// TIA Portal V20 export
// export: Created 2026-10-20T12:39:30.7163103Z, ExportSetting WithDefaults, DisplayName Totally Integrated Automation Portal, DisplayVersion V20 Update 6, DisplayName TIA Portal Openness, DisplayVersion V20 Update 6, DisplayName TIA Portal Version Control Interface, DisplayVersion V20 Update 6, DisplayName SINAMICS Startdrive Advanced, DisplayVersion V20 SP1, DisplayName SINAMICS Startdrive G130, G150, S120, S150, SINAMICS MV, G220, S200, S210, DisplayVersion V20 SP1, DisplayName SINAMICS Startdrive G110M, G120, G120C, G120D, G120P, G115D, DisplayVersion V20 SP1, DisplayName STEP 7 Professional, DisplayVersion V20 Update 6, DisplayName STEP 7 Safety, DisplayVersion V20 Update 2, DisplayName WinCC Basic/Comfort/Advanced, DisplayVersion V20 Update 6, DisplayName WinCC Unified, DisplayVersion V20 Update 6
ORGANIZATION_BLOCK "Main"   // OB1, LAD, ProgramCycle
TITLE = "Main Program Sweep (Cycle)"
{ S7_Optimized_Access := 'TRUE' }
VERSION : 0.1
// stored: AutoNumber true, IsIECCheckEnabled false, SetENOAutomatically false
   VAR_INPUT
      Initial_Call : Bool;   // Initial call of this OB
      Remanence : Bool;   // =True, if remanent data are available
   END_VAR
   VAR_TEMP
      Fault_Handshake_Infeed_1 : Bool;
      Fault_Handshake_Outfeed_1 : Bool;
      Fault_Handshake_Infeed_2 : Bool;
      Fault_Handshake_Infeed_3 : Bool;
      Fault_Handshake_Outfeed_2 : Bool;
      Fault_Handshake_Outfeed_3 : Bool;
   END_VAR
   VAR_TEMP   // added for the SCL form of the ladder/FBD networks
      _w1 : Bool;
      _w2 : Bool;
      _w3 : Bool;
      _w4 : Bool;
      _w5 : Bool;
      _w6 : Bool;
      _w7 : Bool;
      _w8 : Bool;
      _w9 : Bool;
      _w10 : Bool;
      _w11 : Bool;
      _w12 : Bool;
      _w13 : Bool;
      _w14 : Bool;
      _w15 : Bool;
   END_VAR
BEGIN

REGION Network 1: START PLC
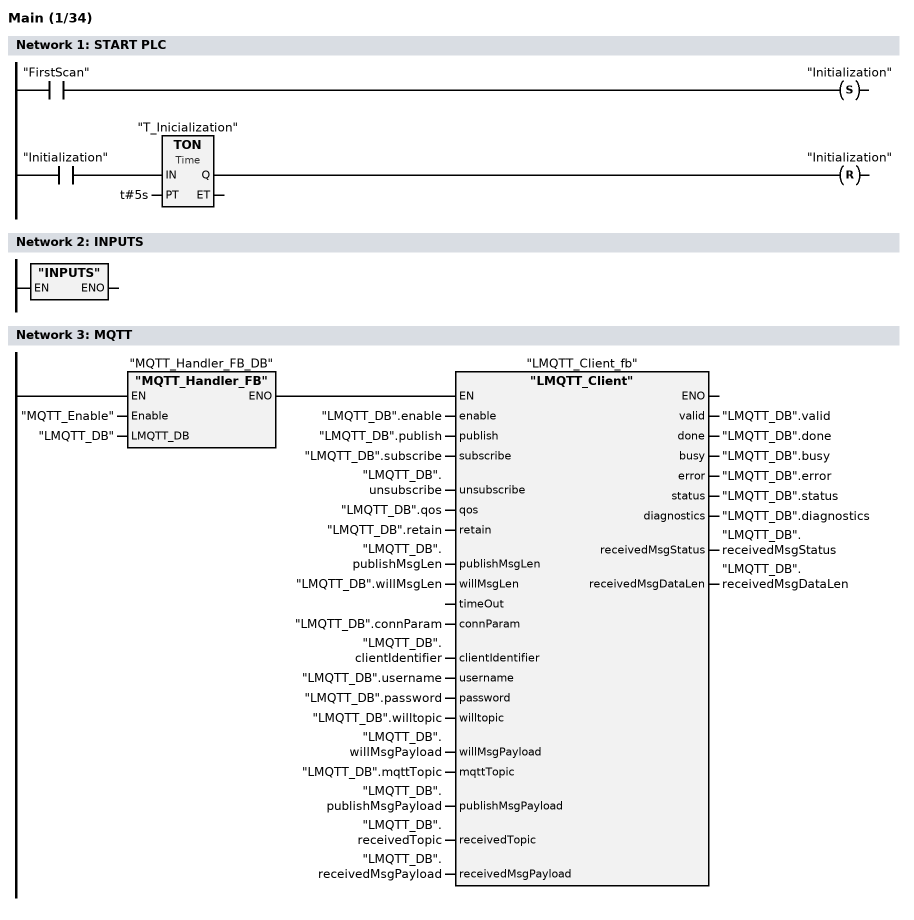
   RUNG wire#powerrail
      Contact( "FirstScan" )
      S_Coil( "Initialization" )
   END_RUNG
   RUNG wire#powerrail
      Contact( "Initialization" )
      { S7_Templates := "time_type := Time" } "T_Inicialization".TON(pt := t#5s, et =>)
      R_Coil( "Initialization" )
   END_RUNG
   // the same network as SCL:
   IF "FirstScan" THEN "Initialization" := TRUE; END_IF;
   "T_Inicialization".TON(IN := "Initialization", PT := t#5s);
   IF "T_Inicialization".Q THEN "Initialization" := FALSE; END_IF;
END_REGION

REGION Network 2: INPUTS
   RUNG wire#powerrail
      "INPUTS"()
   END_RUNG
   // the same network as SCL:
   "INPUTS"();
END_REGION

REGION Network 3: MQTT
   RUNG wire#powerrail
      "MQTT_Handler_FB_DB"(Enable := "MQTT_Enable", LMQTT_DB := "LMQTT_DB")
      "LMQTT_Client_fb"(enable := "LMQTT_DB".enable, publish := "LMQTT_DB".publish, subscribe := "LMQTT_DB".subscribe, unsubscribe := "LMQTT_DB".unsubscribe, qos := "LMQTT_DB".qos, retain := "LMQTT_DB".retain, publishMsgLen := "LMQTT_DB".publishMsgLen, willMsgLen := "LMQTT_DB".willMsgLen, timeOut :=, connParam := "LMQTT_DB".connParam, clientIdentifier := "LMQTT_DB".clientIdentifier, username := "LMQTT_DB".username, password := "LMQTT_DB".password, willtopic := "LMQTT_DB".willtopic, willMsgPayload := "LMQTT_DB".willMsgPayload, mqttTopic := "LMQTT_DB".mqttTopic, publishMsgPayload := "LMQTT_DB".publishMsgPayload, receivedTopic := "LMQTT_DB".receivedTopic, receivedMsgPayload := "LMQTT_DB".receivedMsgPayload, valid => "LMQTT_DB".valid, done => "LMQTT_DB".done, busy => "LMQTT_DB".busy, error => "LMQTT_DB".error, status => "LMQTT_DB".status, diagnostics => "LMQTT_DB".diagnostics, receivedMsgStatus => "LMQTT_DB".receivedMsgStatus, receivedMsgDataLen => "LMQTT_DB".receivedMsgDataLen)
   END_RUNG
   // the same network as SCL:
   "MQTT_Handler_FB_DB"(Enable := "MQTT_Enable", LMQTT_DB := "LMQTT_DB", ENO => #_w1);   // "MQTT_Handler_FB"
   IF #_w1 THEN
       "LMQTT_Client_fb"(enable := "LMQTT_DB".enable,   // "LMQTT_Client"
                         publish := "LMQTT_DB".publish,
                         subscribe := "LMQTT_DB".subscribe,
                         unsubscribe := "LMQTT_DB".unsubscribe,
                         qos := "LMQTT_DB".qos,
                         retain := "LMQTT_DB".retain,
                         publishMsgLen := "LMQTT_DB".publishMsgLen,
                         willMsgLen := "LMQTT_DB".willMsgLen,
                         connParam := "LMQTT_DB".connParam,
                         clientIdentifier := "LMQTT_DB".clientIdentifier,
                         username := "LMQTT_DB".username,
                         password := "LMQTT_DB".password,
                         willtopic := "LMQTT_DB".willtopic,
                         willMsgPayload := "LMQTT_DB".willMsgPayload,
                         mqttTopic := "LMQTT_DB".mqttTopic,
                         publishMsgPayload := "LMQTT_DB".publishMsgPayload,
                         receivedTopic := "LMQTT_DB".receivedTopic,
                         receivedMsgPayload := "LMQTT_DB".receivedMsgPayload,
                         valid => "LMQTT_DB".valid,
                         done => "LMQTT_DB".done,
                         busy => "LMQTT_DB".busy,
                         error => "LMQTT_DB".error,
                         status => "LMQTT_DB".status,
                         diagnostics => "LMQTT_DB".diagnostics,
                         receivedMsgStatus => "LMQTT_DB".receivedMsgStatus,
                         receivedMsgDataLen => "LMQTT_DB".receivedMsgDataLen);
   END_IF;
END_REGION

REGION Network 4: Absolute Encoders
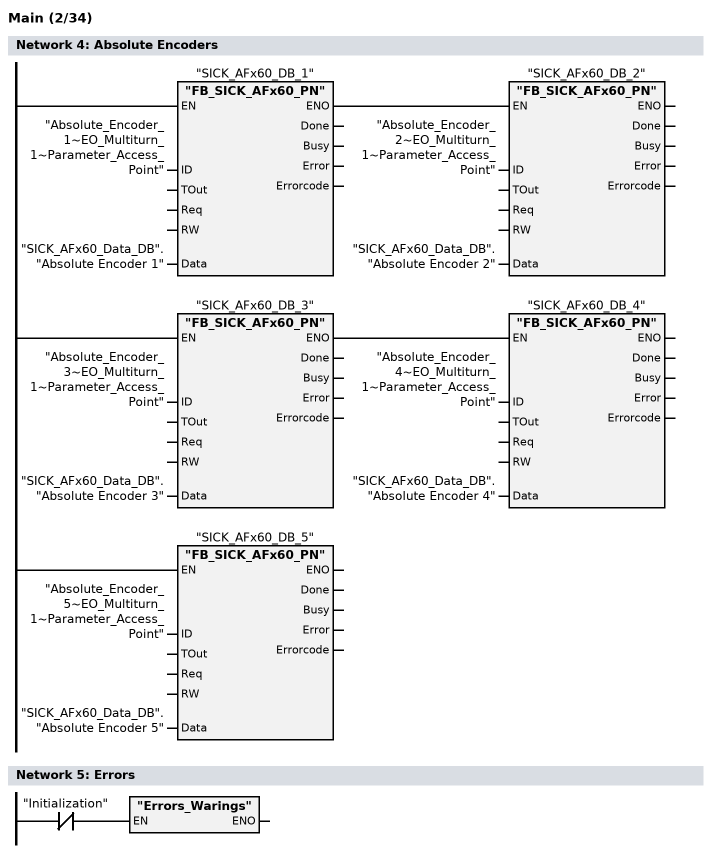
   RUNG wire#powerrail
      "SICK_AFx60_DB_1"(ID := "Absolute_Encoder_1~EO_Multiturn_1~Parameter_Access_Point", TOut :=, Req :=, RW :=, Data := "SICK_AFx60_Data_DB"."Absolute Encoder 1", Done =>, Busy =>, Error =>, Errorcode =>)
      "SICK_AFx60_DB_2"(ID := "Absolute_Encoder_2~EO_Multiturn_1~Parameter_Access_Point", TOut :=, Req :=, RW :=, Data := "SICK_AFx60_Data_DB"."Absolute Encoder 2", Done =>, Busy =>, Error =>, Errorcode =>)
   END_RUNG
   RUNG wire#powerrail
      "SICK_AFx60_DB_3"(ID := "Absolute_Encoder_3~EO_Multiturn_1~Parameter_Access_Point", TOut :=, Req :=, RW :=, Data := "SICK_AFx60_Data_DB"."Absolute Encoder 3", Done =>, Busy =>, Error =>, Errorcode =>)
      "SICK_AFx60_DB_4"(ID := "Absolute_Encoder_4~EO_Multiturn_1~Parameter_Access_Point", TOut :=, Req :=, RW :=, Data := "SICK_AFx60_Data_DB"."Absolute Encoder 4", Done =>, Busy =>, Error =>, Errorcode =>)
   END_RUNG
   RUNG wire#powerrail
      "SICK_AFx60_DB_5"(ID := "Absolute_Encoder_5~EO_Multiturn_1~Parameter_Access_Point", TOut :=, Req :=, RW :=, Data := "SICK_AFx60_Data_DB"."Absolute Encoder 5", Done =>, Busy =>, Error =>, Errorcode =>)
   END_RUNG
   // the same network as SCL:
   "SICK_AFx60_DB_1"(ID := "Absolute_Encoder_1~EO_Multiturn_1~Parameter_Access_Point",   // "FB_SICK_AFx60_PN"
                     Data := "SICK_AFx60_Data_DB"."Absolute Encoder 1",
                     ENO => #_w1);
   IF #_w1 THEN
       "SICK_AFx60_DB_2"(ID := "Absolute_Encoder_2~EO_Multiturn_1~Parameter_Access_Point",   // "FB_SICK_AFx60_PN"
                         Data := "SICK_AFx60_Data_DB"."Absolute Encoder 2");
   END_IF;
   "SICK_AFx60_DB_3"(ID := "Absolute_Encoder_3~EO_Multiturn_1~Parameter_Access_Point",   // "FB_SICK_AFx60_PN"
                     Data := "SICK_AFx60_Data_DB"."Absolute Encoder 3",
                     ENO => #_w2);
   IF #_w2 THEN
       "SICK_AFx60_DB_4"(ID := "Absolute_Encoder_4~EO_Multiturn_1~Parameter_Access_Point",   // "FB_SICK_AFx60_PN"
                         Data := "SICK_AFx60_Data_DB"."Absolute Encoder 4");
   END_IF;
   "SICK_AFx60_DB_5"(ID := "Absolute_Encoder_5~EO_Multiturn_1~Parameter_Access_Point",   // "FB_SICK_AFx60_PN"
                     Data := "SICK_AFx60_Data_DB"."Absolute Encoder 5");
END_REGION

REGION Network 5: Errors
   RUNG wire#powerrail
      I_Contact( "Initialization" )
      "Errors_Warings"()
   END_RUNG
   // the same network as SCL:
   IF NOT "Initialization" THEN "Errors_Warings"(); END_IF;
END_REGION

REGION Network 6: AUTO TEST 1
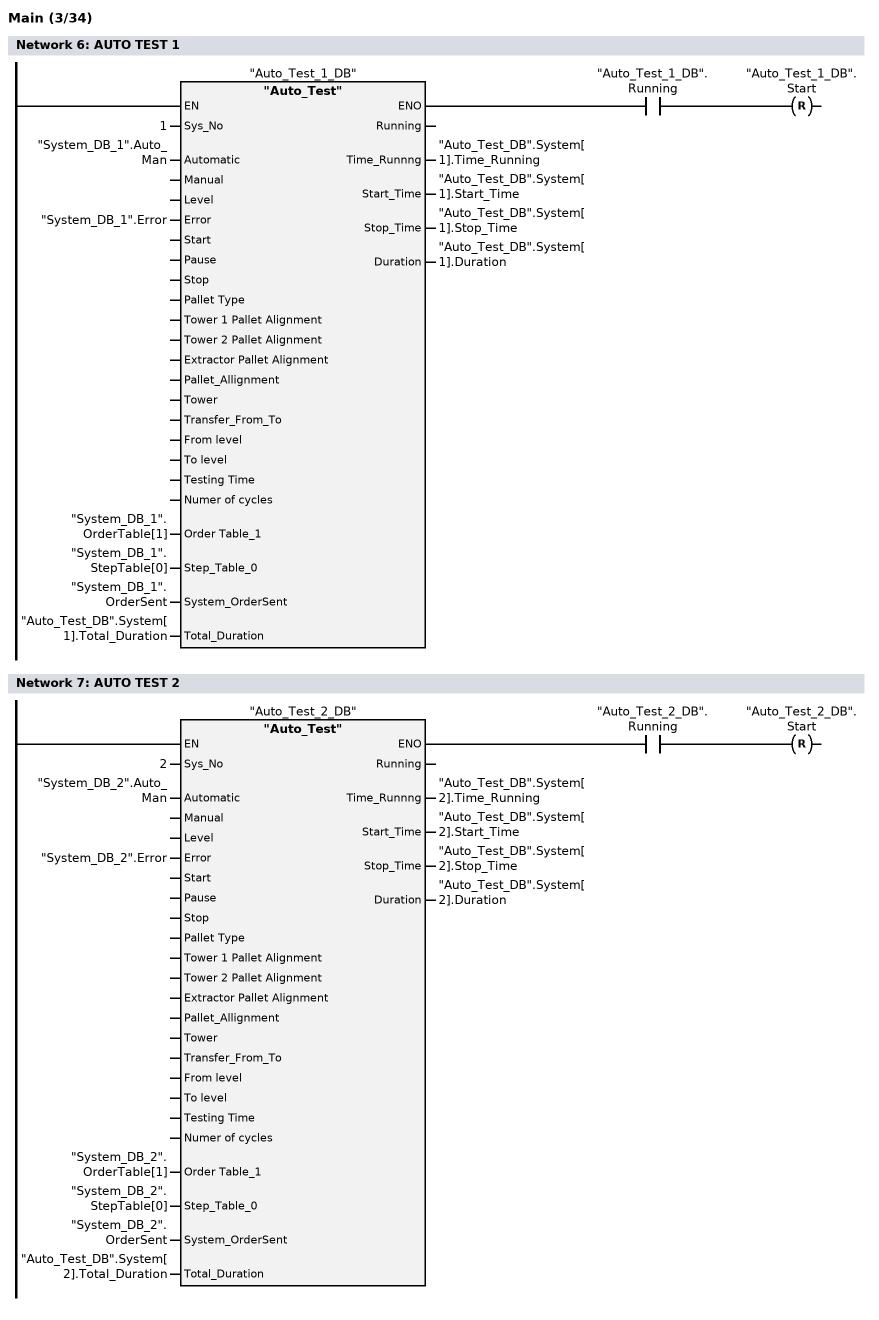
   RUNG wire#powerrail
      "Auto_Test_1_DB"(Sys_No := 1, Automatic := "System_DB_1".Auto_Man, Manual :=, Level :=, Error := "System_DB_1".Error, Start :=, Pause :=, Stop :=, "Pallet Type" :=, "Tower 1 Pallet Alignment" :=, "Tower 2 Pallet Alignment" :=, "Extractor Pallet Alignment" :=, Pallet_Allignment :=, Tower :=, Transfer_From_To :=, "From level" :=, "To level" :=, "Testing Time" :=, "Numer of cycles" :=, "Order Table_1" := "System_DB_1".OrderTable[1], Step_Table_0 := "System_DB_1".StepTable[0], System_OrderSent := "System_DB_1".OrderSent, Total_Duration := "Auto_Test_DB".System[1].Total_Duration, Running =>, Time_Runnng => "Auto_Test_DB".System[1].Time_Running, Start_Time => "Auto_Test_DB".System[1].Start_Time, Stop_Time => "Auto_Test_DB".System[1].Stop_Time, Duration => "Auto_Test_DB".System[1].Duration)
      Contact( "Auto_Test_1_DB".Running )
      R_Coil( "Auto_Test_1_DB".Start )
   END_RUNG
   // the same network as SCL:
   "Auto_Test_1_DB"(Sys_No := 1,   // "Auto_Test"
                    Automatic := "System_DB_1".Auto_Man,
                    Error := "System_DB_1".Error,
                    "Order Table_1" := "System_DB_1".OrderTable[1],
                    Step_Table_0 := "System_DB_1".StepTable[0],
                    System_OrderSent := "System_DB_1".OrderSent,
                    Total_Duration := "Auto_Test_DB".System[1].Total_Duration,
                    Time_Runnng => "Auto_Test_DB".System[1].Time_Running,
                    Start_Time => "Auto_Test_DB".System[1].Start_Time,
                    Stop_Time => "Auto_Test_DB".System[1].Stop_Time,
                    Duration => "Auto_Test_DB".System[1].Duration,
                    ENO => #_w1);
   IF #_w1 AND "Auto_Test_1_DB".Running THEN "Auto_Test_1_DB".Start := FALSE; END_IF;
END_REGION

REGION Network 7: AUTO TEST 2
   RUNG wire#powerrail
      "Auto_Test_2_DB"(Sys_No := 2, Automatic := "System_DB_2".Auto_Man, Manual :=, Level :=, Error := "System_DB_2".Error, Start :=, Pause :=, Stop :=, "Pallet Type" :=, "Tower 1 Pallet Alignment" :=, "Tower 2 Pallet Alignment" :=, "Extractor Pallet Alignment" :=, Pallet_Allignment :=, Tower :=, Transfer_From_To :=, "From level" :=, "To level" :=, "Testing Time" :=, "Numer of cycles" :=, "Order Table_1" := "System_DB_2".OrderTable[1], Step_Table_0 := "System_DB_2".StepTable[0], System_OrderSent := "System_DB_2".OrderSent, Total_Duration := "Auto_Test_DB".System[2].Total_Duration, Running =>, Time_Runnng => "Auto_Test_DB".System[2].Time_Running, Start_Time => "Auto_Test_DB".System[2].Start_Time, Stop_Time => "Auto_Test_DB".System[2].Stop_Time, Duration => "Auto_Test_DB".System[2].Duration)
      Contact( "Auto_Test_2_DB".Running )
      R_Coil( "Auto_Test_2_DB".Start )
   END_RUNG
   // the same network as SCL:
   "Auto_Test_2_DB"(Sys_No := 2,   // "Auto_Test"
                    Automatic := "System_DB_2".Auto_Man,
                    Error := "System_DB_2".Error,
                    "Order Table_1" := "System_DB_2".OrderTable[1],
                    Step_Table_0 := "System_DB_2".StepTable[0],
                    System_OrderSent := "System_DB_2".OrderSent,
                    Total_Duration := "Auto_Test_DB".System[2].Total_Duration,
                    Time_Runnng => "Auto_Test_DB".System[2].Time_Running,
                    Start_Time => "Auto_Test_DB".System[2].Start_Time,
                    Stop_Time => "Auto_Test_DB".System[2].Stop_Time,
                    Duration => "Auto_Test_DB".System[2].Duration,
                    ENO => #_w1);
   IF #_w1 AND "Auto_Test_2_DB".Running THEN "Auto_Test_2_DB".Start := FALSE; END_IF;
END_REGION

REGION Network 8: AUTO TEST 3
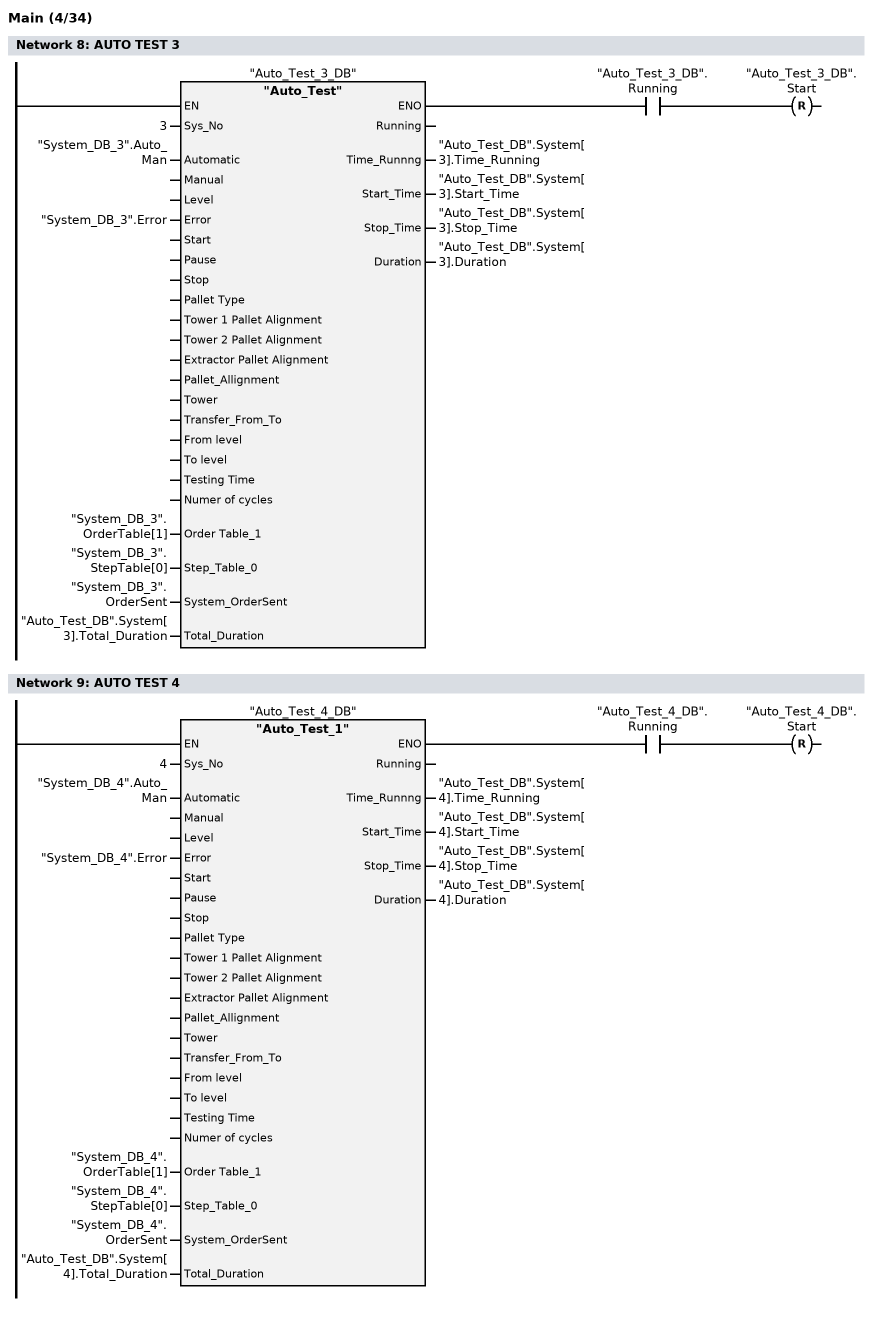
   RUNG wire#powerrail
      "Auto_Test_3_DB"(Sys_No := 3, Automatic := "System_DB_3".Auto_Man, Manual :=, Level :=, Error := "System_DB_3".Error, Start :=, Pause :=, Stop :=, "Pallet Type" :=, "Tower 1 Pallet Alignment" :=, "Tower 2 Pallet Alignment" :=, "Extractor Pallet Alignment" :=, Pallet_Allignment :=, Tower :=, Transfer_From_To :=, "From level" :=, "To level" :=, "Testing Time" :=, "Numer of cycles" :=, "Order Table_1" := "System_DB_3".OrderTable[1], Step_Table_0 := "System_DB_3".StepTable[0], System_OrderSent := "System_DB_3".OrderSent, Total_Duration := "Auto_Test_DB".System[3].Total_Duration, Running =>, Time_Runnng => "Auto_Test_DB".System[3].Time_Running, Start_Time => "Auto_Test_DB".System[3].Start_Time, Stop_Time => "Auto_Test_DB".System[3].Stop_Time, Duration => "Auto_Test_DB".System[3].Duration)
      Contact( "Auto_Test_3_DB".Running )
      R_Coil( "Auto_Test_3_DB".Start )
   END_RUNG
   // the same network as SCL:
   "Auto_Test_3_DB"(Sys_No := 3,   // "Auto_Test"
                    Automatic := "System_DB_3".Auto_Man,
                    Error := "System_DB_3".Error,
                    "Order Table_1" := "System_DB_3".OrderTable[1],
                    Step_Table_0 := "System_DB_3".StepTable[0],
                    System_OrderSent := "System_DB_3".OrderSent,
                    Total_Duration := "Auto_Test_DB".System[3].Total_Duration,
                    Time_Runnng => "Auto_Test_DB".System[3].Time_Running,
                    Start_Time => "Auto_Test_DB".System[3].Start_Time,
                    Stop_Time => "Auto_Test_DB".System[3].Stop_Time,
                    Duration => "Auto_Test_DB".System[3].Duration,
                    ENO => #_w1);
   IF #_w1 AND "Auto_Test_3_DB".Running THEN "Auto_Test_3_DB".Start := FALSE; END_IF;
END_REGION

REGION Network 9: AUTO TEST 4
   RUNG wire#powerrail
      "Auto_Test_4_DB"(Sys_No := 4, Automatic := "System_DB_4".Auto_Man, Manual :=, Level :=, Error := "System_DB_4".Error, Start :=, Pause :=, Stop :=, "Pallet Type" :=, "Tower 1 Pallet Alignment" :=, "Tower 2 Pallet Alignment" :=, "Extractor Pallet Alignment" :=, Pallet_Allignment :=, Tower :=, Transfer_From_To :=, "From level" :=, "To level" :=, "Testing Time" :=, "Numer of cycles" :=, "Order Table_1" := "System_DB_4".OrderTable[1], Step_Table_0 := "System_DB_4".StepTable[0], System_OrderSent := "System_DB_4".OrderSent, Total_Duration := "Auto_Test_DB".System[4].Total_Duration, Running =>, Time_Runnng => "Auto_Test_DB".System[4].Time_Running, Start_Time => "Auto_Test_DB".System[4].Start_Time, Stop_Time => "Auto_Test_DB".System[4].Stop_Time, Duration => "Auto_Test_DB".System[4].Duration)
      Contact( "Auto_Test_4_DB".Running )
      R_Coil( "Auto_Test_4_DB".Start )
   END_RUNG
   // the same network as SCL:
   "Auto_Test_4_DB"(Sys_No := 4,   // "Auto_Test_1"
                    Automatic := "System_DB_4".Auto_Man,
                    Error := "System_DB_4".Error,
                    "Order Table_1" := "System_DB_4".OrderTable[1],
                    Step_Table_0 := "System_DB_4".StepTable[0],
                    System_OrderSent := "System_DB_4".OrderSent,
                    Total_Duration := "Auto_Test_DB".System[4].Total_Duration,
                    Time_Runnng => "Auto_Test_DB".System[4].Time_Running,
                    Start_Time => "Auto_Test_DB".System[4].Start_Time,
                    Stop_Time => "Auto_Test_DB".System[4].Stop_Time,
                    Duration => "Auto_Test_DB".System[4].Duration,
                    ENO => #_w1);
   IF #_w1 AND "Auto_Test_4_DB".Running THEN "Auto_Test_4_DB".Start := FALSE; END_IF;
END_REGION

REGION Network 10: AUTO TEST 5
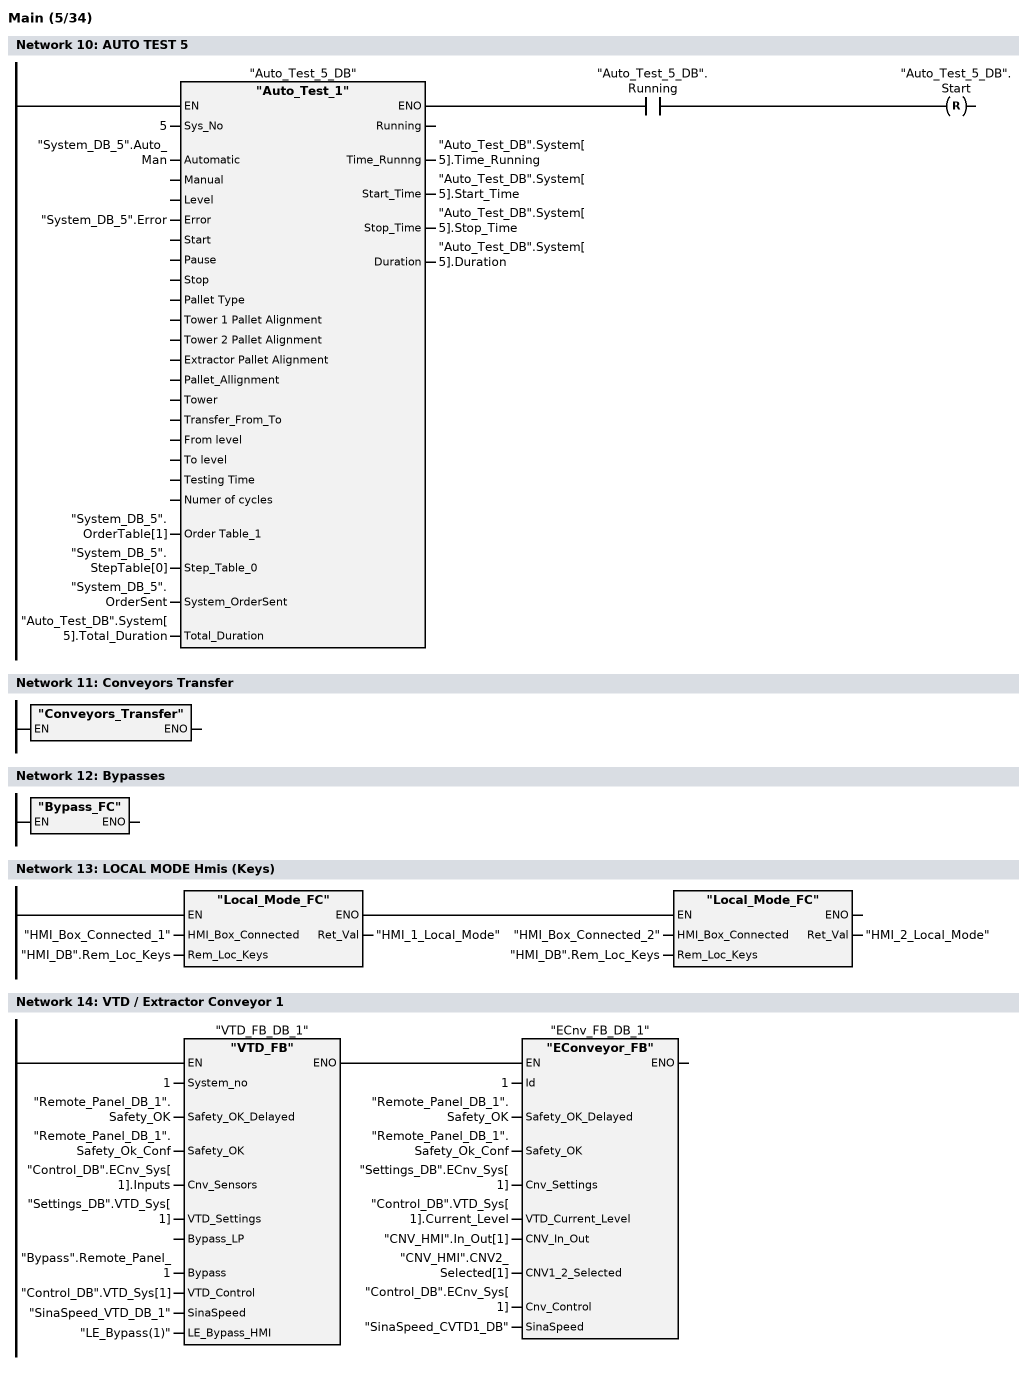
   RUNG wire#powerrail
      "Auto_Test_5_DB"(Sys_No := 5, Automatic := "System_DB_5".Auto_Man, Manual :=, Level :=, Error := "System_DB_5".Error, Start :=, Pause :=, Stop :=, "Pallet Type" :=, "Tower 1 Pallet Alignment" :=, "Tower 2 Pallet Alignment" :=, "Extractor Pallet Alignment" :=, Pallet_Allignment :=, Tower :=, Transfer_From_To :=, "From level" :=, "To level" :=, "Testing Time" :=, "Numer of cycles" :=, "Order Table_1" := "System_DB_5".OrderTable[1], Step_Table_0 := "System_DB_5".StepTable[0], System_OrderSent := "System_DB_5".OrderSent, Total_Duration := "Auto_Test_DB".System[5].Total_Duration, Running =>, Time_Runnng => "Auto_Test_DB".System[5].Time_Running, Start_Time => "Auto_Test_DB".System[5].Start_Time, Stop_Time => "Auto_Test_DB".System[5].Stop_Time, Duration => "Auto_Test_DB".System[5].Duration)
      Contact( "Auto_Test_5_DB".Running )
      R_Coil( "Auto_Test_5_DB".Start )
   END_RUNG
   // the same network as SCL:
   "Auto_Test_5_DB"(Sys_No := 5,   // "Auto_Test_1"
                    Automatic := "System_DB_5".Auto_Man,
                    Error := "System_DB_5".Error,
                    "Order Table_1" := "System_DB_5".OrderTable[1],
                    Step_Table_0 := "System_DB_5".StepTable[0],
                    System_OrderSent := "System_DB_5".OrderSent,
                    Total_Duration := "Auto_Test_DB".System[5].Total_Duration,
                    Time_Runnng => "Auto_Test_DB".System[5].Time_Running,
                    Start_Time => "Auto_Test_DB".System[5].Start_Time,
                    Stop_Time => "Auto_Test_DB".System[5].Stop_Time,
                    Duration => "Auto_Test_DB".System[5].Duration,
                    ENO => #_w1);
   IF #_w1 AND "Auto_Test_5_DB".Running THEN "Auto_Test_5_DB".Start := FALSE; END_IF;
END_REGION

REGION Network 11: Conveyors Transfer
   RUNG wire#powerrail
      "Conveyors_Transfer"()
   END_RUNG
   // the same network as SCL:
   "Conveyors_Transfer"();
END_REGION

REGION Network 12: Bypasses
   RUNG wire#powerrail
      "Bypass_FC"()
   END_RUNG
   // the same network as SCL:
   "Bypass_FC"();
END_REGION

REGION Network 13: LOCAL MODE Hmis (Keys)
   RUNG wire#powerrail
      "Local_Mode_FC"(HMI_Box_Connected := "HMI_Box_Connected_1", Rem_Loc_Keys := "HMI_DB".Rem_Loc_Keys, Ret_Val => "HMI_1_Local_Mode")
      "Local_Mode_FC"(HMI_Box_Connected := "HMI_Box_Connected_2", Rem_Loc_Keys := "HMI_DB".Rem_Loc_Keys, Ret_Val => "HMI_2_Local_Mode")
   END_RUNG
   // the same network as SCL:
   "HMI_1_Local_Mode" := "Local_Mode_FC"(HMI_Box_Connected := "HMI_Box_Connected_1",
                           Rem_Loc_Keys := "HMI_DB".Rem_Loc_Keys,
                           ENO => #_w1);
   IF #_w1 THEN
       "HMI_2_Local_Mode" := "Local_Mode_FC"(HMI_Box_Connected := "HMI_Box_Connected_2",
                               Rem_Loc_Keys := "HMI_DB".Rem_Loc_Keys);
   END_IF;
END_REGION

REGION Network 14: VTD / Extractor Conveyor 1
   RUNG wire#powerrail
      "VTD_FB_DB_1"(System_no := 1, Safety_OK_Delayed := "Remote_Panel_DB_1".Safety_OK, Safety_OK := "Remote_Panel_DB_1".Safety_Ok_Conf, Cnv_Sensors := "Control_DB".ECnv_Sys[1].Inputs, VTD_Settings := "Settings_DB".VTD_Sys[1], Bypass_LP :=, Bypass := "Bypass".Remote_Panel_1, VTD_Control := "Control_DB".VTD_Sys[1], SinaSpeed := "SinaSpeed_VTD_DB_1", LE_Bypass_HMI := "LE_Bypass(1)")
      "ECnv_FB_DB_1"(Id := 1, Safety_OK_Delayed := "Remote_Panel_DB_1".Safety_OK, Safety_OK := "Remote_Panel_DB_1".Safety_Ok_Conf, Cnv_Settings := "Settings_DB".ECnv_Sys[1], VTD_Current_Level := "Control_DB".VTD_Sys[1].Current_Level, CNV_In_Out := "CNV_HMI".In_Out[1], CNV1_2_Selected := "CNV_HMI".CNV2_Selected[1], Cnv_Control := "Control_DB".ECnv_Sys[1], SinaSpeed := "SinaSpeed_CVTD1_DB")
   END_RUNG
   // the same network as SCL:
   "VTD_FB_DB_1"(System_no := 1,   // "VTD_FB"
                 Safety_OK_Delayed := "Remote_Panel_DB_1".Safety_OK,
                 Safety_OK := "Remote_Panel_DB_1".Safety_Ok_Conf,
                 Cnv_Sensors := "Control_DB".ECnv_Sys[1].Inputs,
                 VTD_Settings := "Settings_DB".VTD_Sys[1],
                 Bypass := "Bypass".Remote_Panel_1,
                 VTD_Control := "Control_DB".VTD_Sys[1],
                 SinaSpeed := "SinaSpeed_VTD_DB_1",
                 LE_Bypass_HMI := "LE_Bypass(1)",
                 ENO => #_w1);
   IF #_w1 THEN
       "ECnv_FB_DB_1"(Id := 1,   // "EConveyor_FB"
                      Safety_OK_Delayed := "Remote_Panel_DB_1".Safety_OK,
                      Safety_OK := "Remote_Panel_DB_1".Safety_Ok_Conf,
                      Cnv_Settings := "Settings_DB".ECnv_Sys[1],
                      VTD_Current_Level := "Control_DB".VTD_Sys[1].Current_Level,
                      CNV_In_Out := "CNV_HMI".In_Out[1],
                      CNV1_2_Selected := "CNV_HMI".CNV2_Selected[1],
                      Cnv_Control := "Control_DB".ECnv_Sys[1],
                      SinaSpeed := "SinaSpeed_CVTD1_DB");
   END_IF;
END_REGION

REGION Network 15: VTD / Extractor Conveyor 2
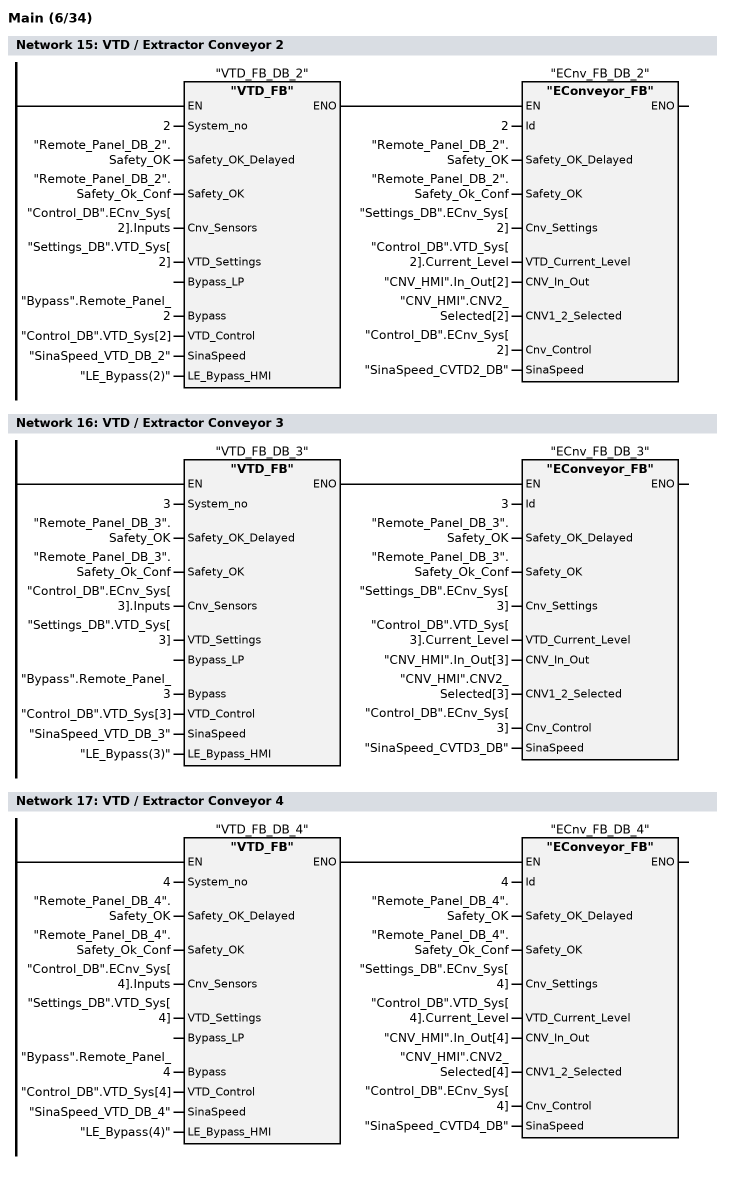
   RUNG wire#powerrail
      "VTD_FB_DB_2"(System_no := 2, Safety_OK_Delayed := "Remote_Panel_DB_2".Safety_OK, Safety_OK := "Remote_Panel_DB_2".Safety_Ok_Conf, Cnv_Sensors := "Control_DB".ECnv_Sys[2].Inputs, VTD_Settings := "Settings_DB".VTD_Sys[2], Bypass_LP :=, Bypass := "Bypass".Remote_Panel_2, VTD_Control := "Control_DB".VTD_Sys[2], SinaSpeed := "SinaSpeed_VTD_DB_2", LE_Bypass_HMI := "LE_Bypass(2)")
      "ECnv_FB_DB_2"(Id := 2, Safety_OK_Delayed := "Remote_Panel_DB_2".Safety_OK, Safety_OK := "Remote_Panel_DB_2".Safety_Ok_Conf, Cnv_Settings := "Settings_DB".ECnv_Sys[2], VTD_Current_Level := "Control_DB".VTD_Sys[2].Current_Level, CNV_In_Out := "CNV_HMI".In_Out[2], CNV1_2_Selected := "CNV_HMI".CNV2_Selected[2], Cnv_Control := "Control_DB".ECnv_Sys[2], SinaSpeed := "SinaSpeed_CVTD2_DB")
   END_RUNG
   // the same network as SCL:
   "VTD_FB_DB_2"(System_no := 2,   // "VTD_FB"
                 Safety_OK_Delayed := "Remote_Panel_DB_2".Safety_OK,
                 Safety_OK := "Remote_Panel_DB_2".Safety_Ok_Conf,
                 Cnv_Sensors := "Control_DB".ECnv_Sys[2].Inputs,
                 VTD_Settings := "Settings_DB".VTD_Sys[2],
                 Bypass := "Bypass".Remote_Panel_2,
                 VTD_Control := "Control_DB".VTD_Sys[2],
                 SinaSpeed := "SinaSpeed_VTD_DB_2",
                 LE_Bypass_HMI := "LE_Bypass(2)",
                 ENO => #_w1);
   IF #_w1 THEN
       "ECnv_FB_DB_2"(Id := 2,   // "EConveyor_FB"
                      Safety_OK_Delayed := "Remote_Panel_DB_2".Safety_OK,
                      Safety_OK := "Remote_Panel_DB_2".Safety_Ok_Conf,
                      Cnv_Settings := "Settings_DB".ECnv_Sys[2],
                      VTD_Current_Level := "Control_DB".VTD_Sys[2].Current_Level,
                      CNV_In_Out := "CNV_HMI".In_Out[2],
                      CNV1_2_Selected := "CNV_HMI".CNV2_Selected[2],
                      Cnv_Control := "Control_DB".ECnv_Sys[2],
                      SinaSpeed := "SinaSpeed_CVTD2_DB");
   END_IF;
END_REGION

REGION Network 16: VTD / Extractor Conveyor 3
   RUNG wire#powerrail
      "VTD_FB_DB_3"(System_no := 3, Safety_OK_Delayed := "Remote_Panel_DB_3".Safety_OK, Safety_OK := "Remote_Panel_DB_3".Safety_Ok_Conf, Cnv_Sensors := "Control_DB".ECnv_Sys[3].Inputs, VTD_Settings := "Settings_DB".VTD_Sys[3], Bypass_LP :=, Bypass := "Bypass".Remote_Panel_3, VTD_Control := "Control_DB".VTD_Sys[3], SinaSpeed := "SinaSpeed_VTD_DB_3", LE_Bypass_HMI := "LE_Bypass(3)")
      "ECnv_FB_DB_3"(Id := 3, Safety_OK_Delayed := "Remote_Panel_DB_3".Safety_OK, Safety_OK := "Remote_Panel_DB_3".Safety_Ok_Conf, Cnv_Settings := "Settings_DB".ECnv_Sys[3], VTD_Current_Level := "Control_DB".VTD_Sys[3].Current_Level, CNV_In_Out := "CNV_HMI".In_Out[3], CNV1_2_Selected := "CNV_HMI".CNV2_Selected[3], Cnv_Control := "Control_DB".ECnv_Sys[3], SinaSpeed := "SinaSpeed_CVTD3_DB")
   END_RUNG
   // the same network as SCL:
   "VTD_FB_DB_3"(System_no := 3,   // "VTD_FB"
                 Safety_OK_Delayed := "Remote_Panel_DB_3".Safety_OK,
                 Safety_OK := "Remote_Panel_DB_3".Safety_Ok_Conf,
                 Cnv_Sensors := "Control_DB".ECnv_Sys[3].Inputs,
                 VTD_Settings := "Settings_DB".VTD_Sys[3],
                 Bypass := "Bypass".Remote_Panel_3,
                 VTD_Control := "Control_DB".VTD_Sys[3],
                 SinaSpeed := "SinaSpeed_VTD_DB_3",
                 LE_Bypass_HMI := "LE_Bypass(3)",
                 ENO => #_w1);
   IF #_w1 THEN
       "ECnv_FB_DB_3"(Id := 3,   // "EConveyor_FB"
                      Safety_OK_Delayed := "Remote_Panel_DB_3".Safety_OK,
                      Safety_OK := "Remote_Panel_DB_3".Safety_Ok_Conf,
                      Cnv_Settings := "Settings_DB".ECnv_Sys[3],
                      VTD_Current_Level := "Control_DB".VTD_Sys[3].Current_Level,
                      CNV_In_Out := "CNV_HMI".In_Out[3],
                      CNV1_2_Selected := "CNV_HMI".CNV2_Selected[3],
                      Cnv_Control := "Control_DB".ECnv_Sys[3],
                      SinaSpeed := "SinaSpeed_CVTD3_DB");
   END_IF;
END_REGION

REGION Network 17: VTD / Extractor Conveyor 4
   RUNG wire#powerrail
      "VTD_FB_DB_4"(System_no := 4, Safety_OK_Delayed := "Remote_Panel_DB_4".Safety_OK, Safety_OK := "Remote_Panel_DB_4".Safety_Ok_Conf, Cnv_Sensors := "Control_DB".ECnv_Sys[4].Inputs, VTD_Settings := "Settings_DB".VTD_Sys[4], Bypass_LP :=, Bypass := "Bypass".Remote_Panel_4, VTD_Control := "Control_DB".VTD_Sys[4], SinaSpeed := "SinaSpeed_VTD_DB_4", LE_Bypass_HMI := "LE_Bypass(4)")
      "ECnv_FB_DB_4"(Id := 4, Safety_OK_Delayed := "Remote_Panel_DB_4".Safety_OK, Safety_OK := "Remote_Panel_DB_4".Safety_Ok_Conf, Cnv_Settings := "Settings_DB".ECnv_Sys[4], VTD_Current_Level := "Control_DB".VTD_Sys[4].Current_Level, CNV_In_Out := "CNV_HMI".In_Out[4], CNV1_2_Selected := "CNV_HMI".CNV2_Selected[4], Cnv_Control := "Control_DB".ECnv_Sys[4], SinaSpeed := "SinaSpeed_CVTD4_DB")
   END_RUNG
   // the same network as SCL:
   "VTD_FB_DB_4"(System_no := 4,   // "VTD_FB"
                 Safety_OK_Delayed := "Remote_Panel_DB_4".Safety_OK,
                 Safety_OK := "Remote_Panel_DB_4".Safety_Ok_Conf,
                 Cnv_Sensors := "Control_DB".ECnv_Sys[4].Inputs,
                 VTD_Settings := "Settings_DB".VTD_Sys[4],
                 Bypass := "Bypass".Remote_Panel_4,
                 VTD_Control := "Control_DB".VTD_Sys[4],
                 SinaSpeed := "SinaSpeed_VTD_DB_4",
                 LE_Bypass_HMI := "LE_Bypass(4)",
                 ENO => #_w1);
   IF #_w1 THEN
       "ECnv_FB_DB_4"(Id := 4,   // "EConveyor_FB"
                      Safety_OK_Delayed := "Remote_Panel_DB_4".Safety_OK,
                      Safety_OK := "Remote_Panel_DB_4".Safety_Ok_Conf,
                      Cnv_Settings := "Settings_DB".ECnv_Sys[4],
                      VTD_Current_Level := "Control_DB".VTD_Sys[4].Current_Level,
                      CNV_In_Out := "CNV_HMI".In_Out[4],
                      CNV1_2_Selected := "CNV_HMI".CNV2_Selected[4],
                      Cnv_Control := "Control_DB".ECnv_Sys[4],
                      SinaSpeed := "SinaSpeed_CVTD4_DB");
   END_IF;
END_REGION

REGION Network 18: VTD / Extractor Conveyor 5
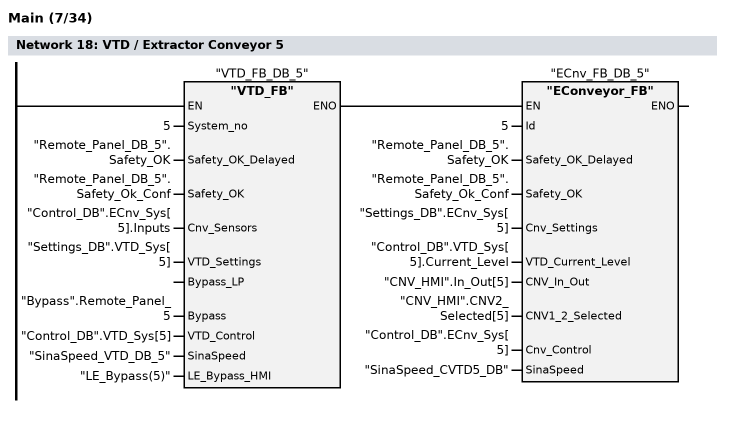
   RUNG wire#powerrail
      "VTD_FB_DB_5"(System_no := 5, Safety_OK_Delayed := "Remote_Panel_DB_5".Safety_OK, Safety_OK := "Remote_Panel_DB_5".Safety_Ok_Conf, Cnv_Sensors := "Control_DB".ECnv_Sys[5].Inputs, VTD_Settings := "Settings_DB".VTD_Sys[5], Bypass_LP :=, Bypass := "Bypass".Remote_Panel_5, VTD_Control := "Control_DB".VTD_Sys[5], SinaSpeed := "SinaSpeed_VTD_DB_5", LE_Bypass_HMI := "LE_Bypass(5)")
      "ECnv_FB_DB_5"(Id := 5, Safety_OK_Delayed := "Remote_Panel_DB_5".Safety_OK, Safety_OK := "Remote_Panel_DB_5".Safety_Ok_Conf, Cnv_Settings := "Settings_DB".ECnv_Sys[5], VTD_Current_Level := "Control_DB".VTD_Sys[5].Current_Level, CNV_In_Out := "CNV_HMI".In_Out[5], CNV1_2_Selected := "CNV_HMI".CNV2_Selected[5], Cnv_Control := "Control_DB".ECnv_Sys[5], SinaSpeed := "SinaSpeed_CVTD5_DB")
   END_RUNG
   // the same network as SCL:
   "VTD_FB_DB_5"(System_no := 5,   // "VTD_FB"
                 Safety_OK_Delayed := "Remote_Panel_DB_5".Safety_OK,
                 Safety_OK := "Remote_Panel_DB_5".Safety_Ok_Conf,
                 Cnv_Sensors := "Control_DB".ECnv_Sys[5].Inputs,
                 VTD_Settings := "Settings_DB".VTD_Sys[5],
                 Bypass := "Bypass".Remote_Panel_5,
                 VTD_Control := "Control_DB".VTD_Sys[5],
                 SinaSpeed := "SinaSpeed_VTD_DB_5",
                 LE_Bypass_HMI := "LE_Bypass(5)",
                 ENO => #_w1);
   IF #_w1 THEN
       "ECnv_FB_DB_5"(Id := 5,   // "EConveyor_FB"
                      Safety_OK_Delayed := "Remote_Panel_DB_5".Safety_OK,
                      Safety_OK := "Remote_Panel_DB_5".Safety_Ok_Conf,
                      Cnv_Settings := "Settings_DB".ECnv_Sys[5],
                      VTD_Current_Level := "Control_DB".VTD_Sys[5].Current_Level,
                      CNV_In_Out := "CNV_HMI".In_Out[5],
                      CNV1_2_Selected := "CNV_HMI".CNV2_Selected[5],
                      Cnv_Control := "Control_DB".ECnv_Sys[5],
                      SinaSpeed := "SinaSpeed_CVTD5_DB");
   END_IF;
END_REGION

REGION Network 19: SYSTEM 1
END_REGION

REGION Network 20: Level Conveyors Tower 1 - SYSTEM 1
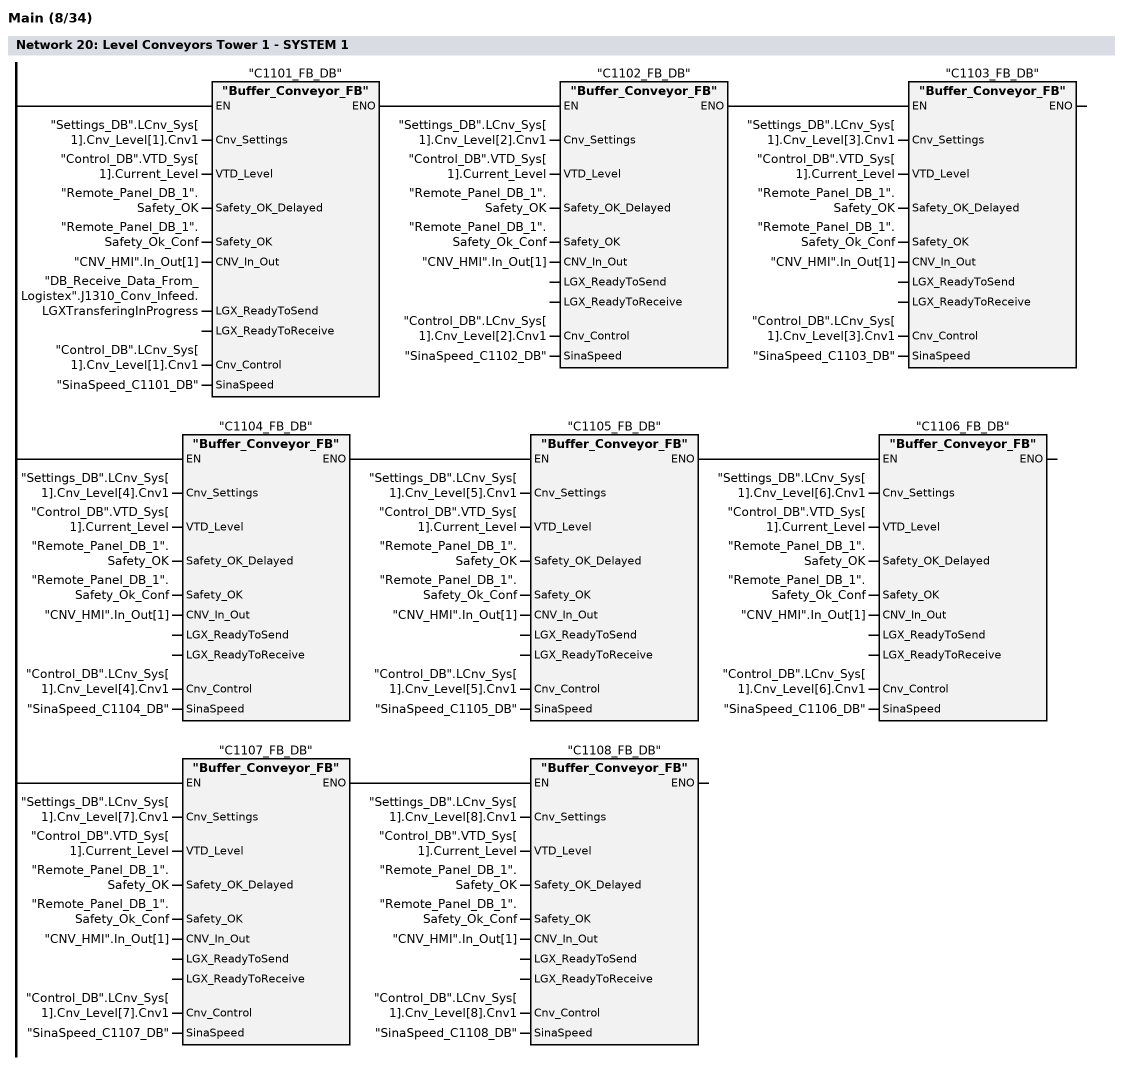
   RUNG wire#powerrail
      "C1101_FB_DB"(Cnv_Settings := "Settings_DB".LCnv_Sys[1].Cnv_Level[1].Cnv1, VTD_Level := "Control_DB".VTD_Sys[1].Current_Level, Safety_OK_Delayed := "Remote_Panel_DB_1".Safety_OK, Safety_OK := "Remote_Panel_DB_1".Safety_Ok_Conf, CNV_In_Out := "CNV_HMI".In_Out[1], LGX_ReadyToSend := "DB_Receive_Data_From_Logistex".J1310_Conv_Infeed.LGXTransferingInProgress, LGX_ReadyToReceive :=, Cnv_Control := "Control_DB".LCnv_Sys[1].Cnv_Level[1].Cnv1, SinaSpeed := "SinaSpeed_C1101_DB")
      "C1102_FB_DB"(Cnv_Settings := "Settings_DB".LCnv_Sys[1].Cnv_Level[2].Cnv1, VTD_Level := "Control_DB".VTD_Sys[1].Current_Level, Safety_OK_Delayed := "Remote_Panel_DB_1".Safety_OK, Safety_OK := "Remote_Panel_DB_1".Safety_Ok_Conf, CNV_In_Out := "CNV_HMI".In_Out[1], LGX_ReadyToSend :=, LGX_ReadyToReceive :=, Cnv_Control := "Control_DB".LCnv_Sys[1].Cnv_Level[2].Cnv1, SinaSpeed := "SinaSpeed_C1102_DB")
      "C1103_FB_DB"(Cnv_Settings := "Settings_DB".LCnv_Sys[1].Cnv_Level[3].Cnv1, VTD_Level := "Control_DB".VTD_Sys[1].Current_Level, Safety_OK_Delayed := "Remote_Panel_DB_1".Safety_OK, Safety_OK := "Remote_Panel_DB_1".Safety_Ok_Conf, CNV_In_Out := "CNV_HMI".In_Out[1], LGX_ReadyToSend :=, LGX_ReadyToReceive :=, Cnv_Control := "Control_DB".LCnv_Sys[1].Cnv_Level[3].Cnv1, SinaSpeed := "SinaSpeed_C1103_DB")
   END_RUNG
   RUNG wire#powerrail
      "C1104_FB_DB"(Cnv_Settings := "Settings_DB".LCnv_Sys[1].Cnv_Level[4].Cnv1, VTD_Level := "Control_DB".VTD_Sys[1].Current_Level, Safety_OK_Delayed := "Remote_Panel_DB_1".Safety_OK, Safety_OK := "Remote_Panel_DB_1".Safety_Ok_Conf, CNV_In_Out := "CNV_HMI".In_Out[1], LGX_ReadyToSend :=, LGX_ReadyToReceive :=, Cnv_Control := "Control_DB".LCnv_Sys[1].Cnv_Level[4].Cnv1, SinaSpeed := "SinaSpeed_C1104_DB")
      "C1105_FB_DB"(Cnv_Settings := "Settings_DB".LCnv_Sys[1].Cnv_Level[5].Cnv1, VTD_Level := "Control_DB".VTD_Sys[1].Current_Level, Safety_OK_Delayed := "Remote_Panel_DB_1".Safety_OK, Safety_OK := "Remote_Panel_DB_1".Safety_Ok_Conf, CNV_In_Out := "CNV_HMI".In_Out[1], LGX_ReadyToSend :=, LGX_ReadyToReceive :=, Cnv_Control := "Control_DB".LCnv_Sys[1].Cnv_Level[5].Cnv1, SinaSpeed := "SinaSpeed_C1105_DB")
      "C1106_FB_DB"(Cnv_Settings := "Settings_DB".LCnv_Sys[1].Cnv_Level[6].Cnv1, VTD_Level := "Control_DB".VTD_Sys[1].Current_Level, Safety_OK_Delayed := "Remote_Panel_DB_1".Safety_OK, Safety_OK := "Remote_Panel_DB_1".Safety_Ok_Conf, CNV_In_Out := "CNV_HMI".In_Out[1], LGX_ReadyToSend :=, LGX_ReadyToReceive :=, Cnv_Control := "Control_DB".LCnv_Sys[1].Cnv_Level[6].Cnv1, SinaSpeed := "SinaSpeed_C1106_DB")
   END_RUNG
   RUNG wire#powerrail
      "C1107_FB_DB"(Cnv_Settings := "Settings_DB".LCnv_Sys[1].Cnv_Level[7].Cnv1, VTD_Level := "Control_DB".VTD_Sys[1].Current_Level, Safety_OK_Delayed := "Remote_Panel_DB_1".Safety_OK, Safety_OK := "Remote_Panel_DB_1".Safety_Ok_Conf, CNV_In_Out := "CNV_HMI".In_Out[1], LGX_ReadyToSend :=, LGX_ReadyToReceive :=, Cnv_Control := "Control_DB".LCnv_Sys[1].Cnv_Level[7].Cnv1, SinaSpeed := "SinaSpeed_C1107_DB")
      "C1108_FB_DB"(Cnv_Settings := "Settings_DB".LCnv_Sys[1].Cnv_Level[8].Cnv1, VTD_Level := "Control_DB".VTD_Sys[1].Current_Level, Safety_OK_Delayed := "Remote_Panel_DB_1".Safety_OK, Safety_OK := "Remote_Panel_DB_1".Safety_Ok_Conf, CNV_In_Out := "CNV_HMI".In_Out[1], LGX_ReadyToSend :=, LGX_ReadyToReceive :=, Cnv_Control := "Control_DB".LCnv_Sys[1].Cnv_Level[8].Cnv1, SinaSpeed := "SinaSpeed_C1108_DB")
   END_RUNG
   // the same network as SCL:
   "C1101_FB_DB"(Cnv_Settings := "Settings_DB".LCnv_Sys[1].Cnv_Level[1].Cnv1,   // "Buffer_Conveyor_FB"
                 VTD_Level := "Control_DB".VTD_Sys[1].Current_Level,
                 Safety_OK_Delayed := "Remote_Panel_DB_1".Safety_OK,
                 Safety_OK := "Remote_Panel_DB_1".Safety_Ok_Conf,
                 CNV_In_Out := "CNV_HMI".In_Out[1],
                 LGX_ReadyToSend := "DB_Receive_Data_From_Logistex".J1310_Conv_Infeed.LGXTransferingInProgress,
                 Cnv_Control := "Control_DB".LCnv_Sys[1].Cnv_Level[1].Cnv1,
                 SinaSpeed := "SinaSpeed_C1101_DB",
                 ENO => #_w1);
   "C1102_FB_DB"(EN := #_w1,   // "Buffer_Conveyor_FB"
                 Cnv_Settings := "Settings_DB".LCnv_Sys[1].Cnv_Level[2].Cnv1,
                 VTD_Level := "Control_DB".VTD_Sys[1].Current_Level,
                 Safety_OK_Delayed := "Remote_Panel_DB_1".Safety_OK,
                 Safety_OK := "Remote_Panel_DB_1".Safety_Ok_Conf,
                 CNV_In_Out := "CNV_HMI".In_Out[1],
                 Cnv_Control := "Control_DB".LCnv_Sys[1].Cnv_Level[2].Cnv1,
                 SinaSpeed := "SinaSpeed_C1102_DB",
                 ENO => #_w2);
   IF #_w2 THEN
       "C1103_FB_DB"(Cnv_Settings := "Settings_DB".LCnv_Sys[1].Cnv_Level[3].Cnv1,   // "Buffer_Conveyor_FB"
                     VTD_Level := "Control_DB".VTD_Sys[1].Current_Level,
                     Safety_OK_Delayed := "Remote_Panel_DB_1".Safety_OK,
                     Safety_OK := "Remote_Panel_DB_1".Safety_Ok_Conf,
                     CNV_In_Out := "CNV_HMI".In_Out[1],
                     Cnv_Control := "Control_DB".LCnv_Sys[1].Cnv_Level[3].Cnv1,
                     SinaSpeed := "SinaSpeed_C1103_DB");
   END_IF;
   "C1104_FB_DB"(Cnv_Settings := "Settings_DB".LCnv_Sys[1].Cnv_Level[4].Cnv1,   // "Buffer_Conveyor_FB"
                 VTD_Level := "Control_DB".VTD_Sys[1].Current_Level,
                 Safety_OK_Delayed := "Remote_Panel_DB_1".Safety_OK,
                 Safety_OK := "Remote_Panel_DB_1".Safety_Ok_Conf,
                 CNV_In_Out := "CNV_HMI".In_Out[1],
                 Cnv_Control := "Control_DB".LCnv_Sys[1].Cnv_Level[4].Cnv1,
                 SinaSpeed := "SinaSpeed_C1104_DB",
                 ENO => #_w3);
   "C1105_FB_DB"(EN := #_w3,   // "Buffer_Conveyor_FB"
                 Cnv_Settings := "Settings_DB".LCnv_Sys[1].Cnv_Level[5].Cnv1,
                 VTD_Level := "Control_DB".VTD_Sys[1].Current_Level,
                 Safety_OK_Delayed := "Remote_Panel_DB_1".Safety_OK,
                 Safety_OK := "Remote_Panel_DB_1".Safety_Ok_Conf,
                 CNV_In_Out := "CNV_HMI".In_Out[1],
                 Cnv_Control := "Control_DB".LCnv_Sys[1].Cnv_Level[5].Cnv1,
                 SinaSpeed := "SinaSpeed_C1105_DB",
                 ENO => #_w4);
   IF #_w4 THEN
       "C1106_FB_DB"(Cnv_Settings := "Settings_DB".LCnv_Sys[1].Cnv_Level[6].Cnv1,   // "Buffer_Conveyor_FB"
                     VTD_Level := "Control_DB".VTD_Sys[1].Current_Level,
                     Safety_OK_Delayed := "Remote_Panel_DB_1".Safety_OK,
                     Safety_OK := "Remote_Panel_DB_1".Safety_Ok_Conf,
                     CNV_In_Out := "CNV_HMI".In_Out[1],
                     Cnv_Control := "Control_DB".LCnv_Sys[1].Cnv_Level[6].Cnv1,
                     SinaSpeed := "SinaSpeed_C1106_DB");
   END_IF;
   "C1107_FB_DB"(Cnv_Settings := "Settings_DB".LCnv_Sys[1].Cnv_Level[7].Cnv1,   // "Buffer_Conveyor_FB"
                 VTD_Level := "Control_DB".VTD_Sys[1].Current_Level,
                 Safety_OK_Delayed := "Remote_Panel_DB_1".Safety_OK,
                 Safety_OK := "Remote_Panel_DB_1".Safety_Ok_Conf,
                 CNV_In_Out := "CNV_HMI".In_Out[1],
                 Cnv_Control := "Control_DB".LCnv_Sys[1].Cnv_Level[7].Cnv1,
                 SinaSpeed := "SinaSpeed_C1107_DB",
                 ENO => #_w5);
   IF #_w5 THEN
       "C1108_FB_DB"(Cnv_Settings := "Settings_DB".LCnv_Sys[1].Cnv_Level[8].Cnv1,   // "Buffer_Conveyor_FB"
                     VTD_Level := "Control_DB".VTD_Sys[1].Current_Level,
                     Safety_OK_Delayed := "Remote_Panel_DB_1".Safety_OK,
                     Safety_OK := "Remote_Panel_DB_1".Safety_Ok_Conf,
                     CNV_In_Out := "CNV_HMI".In_Out[1],
                     Cnv_Control := "Control_DB".LCnv_Sys[1].Cnv_Level[8].Cnv1,
                     SinaSpeed := "SinaSpeed_C1108_DB");
   END_IF;
END_REGION

REGION Network 21: Level Conveyors Tower 2 - SYSTEM 1
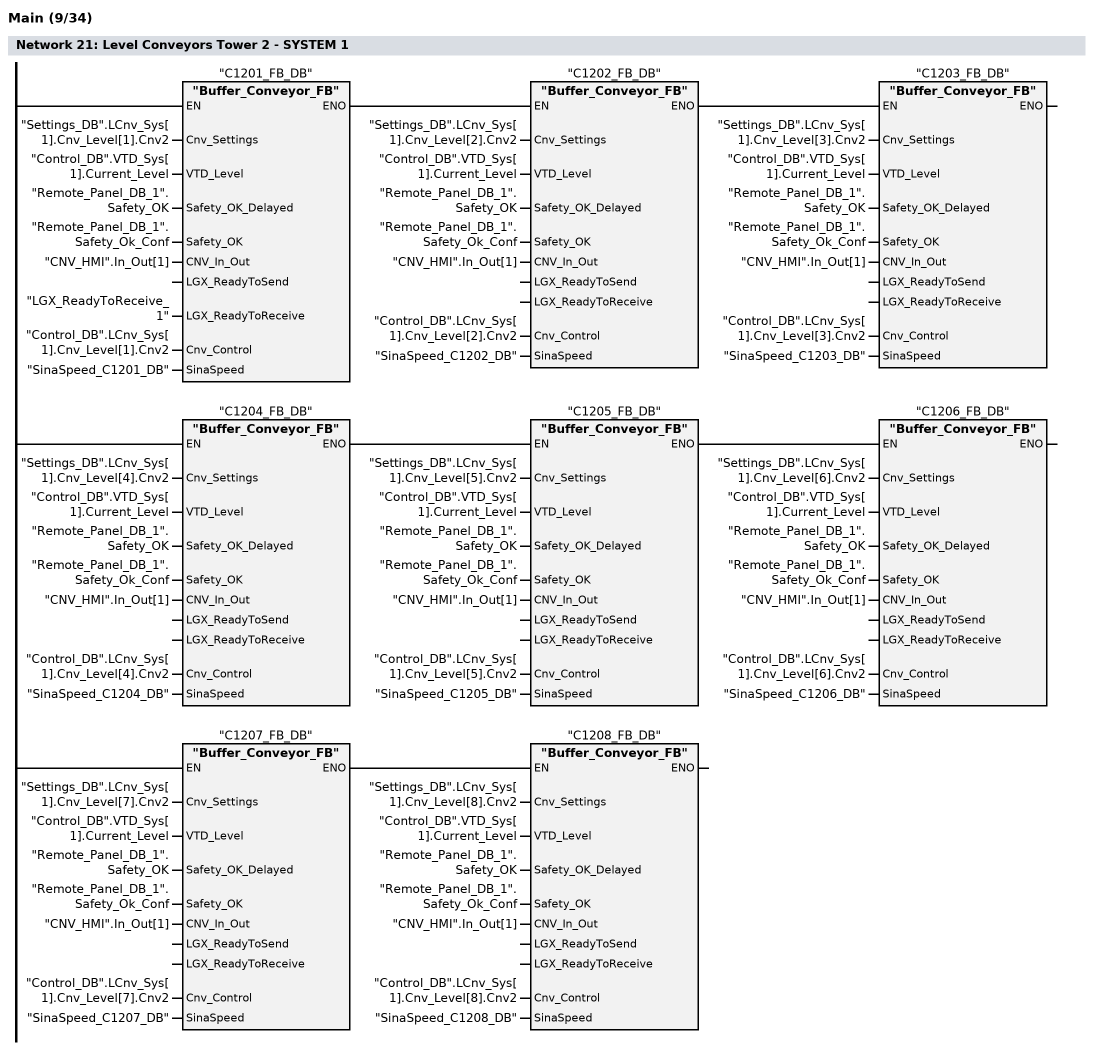
   RUNG wire#powerrail
      "C1201_FB_DB"(Cnv_Settings := "Settings_DB".LCnv_Sys[1].Cnv_Level[1].Cnv2, VTD_Level := "Control_DB".VTD_Sys[1].Current_Level, Safety_OK_Delayed := "Remote_Panel_DB_1".Safety_OK, Safety_OK := "Remote_Panel_DB_1".Safety_Ok_Conf, CNV_In_Out := "CNV_HMI".In_Out[1], LGX_ReadyToSend :=, LGX_ReadyToReceive := "LGX_ReadyToReceive_1", Cnv_Control := "Control_DB".LCnv_Sys[1].Cnv_Level[1].Cnv2, SinaSpeed := "SinaSpeed_C1201_DB")
      "C1202_FB_DB"(Cnv_Settings := "Settings_DB".LCnv_Sys[1].Cnv_Level[2].Cnv2, VTD_Level := "Control_DB".VTD_Sys[1].Current_Level, Safety_OK_Delayed := "Remote_Panel_DB_1".Safety_OK, Safety_OK := "Remote_Panel_DB_1".Safety_Ok_Conf, CNV_In_Out := "CNV_HMI".In_Out[1], LGX_ReadyToSend :=, LGX_ReadyToReceive :=, Cnv_Control := "Control_DB".LCnv_Sys[1].Cnv_Level[2].Cnv2, SinaSpeed := "SinaSpeed_C1202_DB")
      "C1203_FB_DB"(Cnv_Settings := "Settings_DB".LCnv_Sys[1].Cnv_Level[3].Cnv2, VTD_Level := "Control_DB".VTD_Sys[1].Current_Level, Safety_OK_Delayed := "Remote_Panel_DB_1".Safety_OK, Safety_OK := "Remote_Panel_DB_1".Safety_Ok_Conf, CNV_In_Out := "CNV_HMI".In_Out[1], LGX_ReadyToSend :=, LGX_ReadyToReceive :=, Cnv_Control := "Control_DB".LCnv_Sys[1].Cnv_Level[3].Cnv2, SinaSpeed := "SinaSpeed_C1203_DB")
   END_RUNG
   RUNG wire#powerrail
      "C1204_FB_DB"(Cnv_Settings := "Settings_DB".LCnv_Sys[1].Cnv_Level[4].Cnv2, VTD_Level := "Control_DB".VTD_Sys[1].Current_Level, Safety_OK_Delayed := "Remote_Panel_DB_1".Safety_OK, Safety_OK := "Remote_Panel_DB_1".Safety_Ok_Conf, CNV_In_Out := "CNV_HMI".In_Out[1], LGX_ReadyToSend :=, LGX_ReadyToReceive :=, Cnv_Control := "Control_DB".LCnv_Sys[1].Cnv_Level[4].Cnv2, SinaSpeed := "SinaSpeed_C1204_DB")
      "C1205_FB_DB"(Cnv_Settings := "Settings_DB".LCnv_Sys[1].Cnv_Level[5].Cnv2, VTD_Level := "Control_DB".VTD_Sys[1].Current_Level, Safety_OK_Delayed := "Remote_Panel_DB_1".Safety_OK, Safety_OK := "Remote_Panel_DB_1".Safety_Ok_Conf, CNV_In_Out := "CNV_HMI".In_Out[1], LGX_ReadyToSend :=, LGX_ReadyToReceive :=, Cnv_Control := "Control_DB".LCnv_Sys[1].Cnv_Level[5].Cnv2, SinaSpeed := "SinaSpeed_C1205_DB")
      "C1206_FB_DB"(Cnv_Settings := "Settings_DB".LCnv_Sys[1].Cnv_Level[6].Cnv2, VTD_Level := "Control_DB".VTD_Sys[1].Current_Level, Safety_OK_Delayed := "Remote_Panel_DB_1".Safety_OK, Safety_OK := "Remote_Panel_DB_1".Safety_Ok_Conf, CNV_In_Out := "CNV_HMI".In_Out[1], LGX_ReadyToSend :=, LGX_ReadyToReceive :=, Cnv_Control := "Control_DB".LCnv_Sys[1].Cnv_Level[6].Cnv2, SinaSpeed := "SinaSpeed_C1206_DB")
   END_RUNG
   RUNG wire#powerrail
      "C1207_FB_DB"(Cnv_Settings := "Settings_DB".LCnv_Sys[1].Cnv_Level[7].Cnv2, VTD_Level := "Control_DB".VTD_Sys[1].Current_Level, Safety_OK_Delayed := "Remote_Panel_DB_1".Safety_OK, Safety_OK := "Remote_Panel_DB_1".Safety_Ok_Conf, CNV_In_Out := "CNV_HMI".In_Out[1], LGX_ReadyToSend :=, LGX_ReadyToReceive :=, Cnv_Control := "Control_DB".LCnv_Sys[1].Cnv_Level[7].Cnv2, SinaSpeed := "SinaSpeed_C1207_DB")
      "C1208_FB_DB"(Cnv_Settings := "Settings_DB".LCnv_Sys[1].Cnv_Level[8].Cnv2, VTD_Level := "Control_DB".VTD_Sys[1].Current_Level, Safety_OK_Delayed := "Remote_Panel_DB_1".Safety_OK, Safety_OK := "Remote_Panel_DB_1".Safety_Ok_Conf, CNV_In_Out := "CNV_HMI".In_Out[1], LGX_ReadyToSend :=, LGX_ReadyToReceive :=, Cnv_Control := "Control_DB".LCnv_Sys[1].Cnv_Level[8].Cnv2, SinaSpeed := "SinaSpeed_C1208_DB")
   END_RUNG
   // the same network as SCL:
   "C1201_FB_DB"(Cnv_Settings := "Settings_DB".LCnv_Sys[1].Cnv_Level[1].Cnv2,   // "Buffer_Conveyor_FB"
                 VTD_Level := "Control_DB".VTD_Sys[1].Current_Level,
                 Safety_OK_Delayed := "Remote_Panel_DB_1".Safety_OK,
                 Safety_OK := "Remote_Panel_DB_1".Safety_Ok_Conf,
                 CNV_In_Out := "CNV_HMI".In_Out[1],
                 LGX_ReadyToReceive := "LGX_ReadyToReceive_1",
                 Cnv_Control := "Control_DB".LCnv_Sys[1].Cnv_Level[1].Cnv2,
                 SinaSpeed := "SinaSpeed_C1201_DB",
                 ENO => #_w1);
   "C1202_FB_DB"(EN := #_w1,   // "Buffer_Conveyor_FB"
                 Cnv_Settings := "Settings_DB".LCnv_Sys[1].Cnv_Level[2].Cnv2,
                 VTD_Level := "Control_DB".VTD_Sys[1].Current_Level,
                 Safety_OK_Delayed := "Remote_Panel_DB_1".Safety_OK,
                 Safety_OK := "Remote_Panel_DB_1".Safety_Ok_Conf,
                 CNV_In_Out := "CNV_HMI".In_Out[1],
                 Cnv_Control := "Control_DB".LCnv_Sys[1].Cnv_Level[2].Cnv2,
                 SinaSpeed := "SinaSpeed_C1202_DB",
                 ENO => #_w2);
   IF #_w2 THEN
       "C1203_FB_DB"(Cnv_Settings := "Settings_DB".LCnv_Sys[1].Cnv_Level[3].Cnv2,   // "Buffer_Conveyor_FB"
                     VTD_Level := "Control_DB".VTD_Sys[1].Current_Level,
                     Safety_OK_Delayed := "Remote_Panel_DB_1".Safety_OK,
                     Safety_OK := "Remote_Panel_DB_1".Safety_Ok_Conf,
                     CNV_In_Out := "CNV_HMI".In_Out[1],
                     Cnv_Control := "Control_DB".LCnv_Sys[1].Cnv_Level[3].Cnv2,
                     SinaSpeed := "SinaSpeed_C1203_DB");
   END_IF;
   "C1204_FB_DB"(Cnv_Settings := "Settings_DB".LCnv_Sys[1].Cnv_Level[4].Cnv2,   // "Buffer_Conveyor_FB"
                 VTD_Level := "Control_DB".VTD_Sys[1].Current_Level,
                 Safety_OK_Delayed := "Remote_Panel_DB_1".Safety_OK,
                 Safety_OK := "Remote_Panel_DB_1".Safety_Ok_Conf,
                 CNV_In_Out := "CNV_HMI".In_Out[1],
                 Cnv_Control := "Control_DB".LCnv_Sys[1].Cnv_Level[4].Cnv2,
                 SinaSpeed := "SinaSpeed_C1204_DB",
                 ENO => #_w3);
   "C1205_FB_DB"(EN := #_w3,   // "Buffer_Conveyor_FB"
                 Cnv_Settings := "Settings_DB".LCnv_Sys[1].Cnv_Level[5].Cnv2,
                 VTD_Level := "Control_DB".VTD_Sys[1].Current_Level,
                 Safety_OK_Delayed := "Remote_Panel_DB_1".Safety_OK,
                 Safety_OK := "Remote_Panel_DB_1".Safety_Ok_Conf,
                 CNV_In_Out := "CNV_HMI".In_Out[1],
                 Cnv_Control := "Control_DB".LCnv_Sys[1].Cnv_Level[5].Cnv2,
                 SinaSpeed := "SinaSpeed_C1205_DB",
                 ENO => #_w4);
   IF #_w4 THEN
       "C1206_FB_DB"(Cnv_Settings := "Settings_DB".LCnv_Sys[1].Cnv_Level[6].Cnv2,   // "Buffer_Conveyor_FB"
                     VTD_Level := "Control_DB".VTD_Sys[1].Current_Level,
                     Safety_OK_Delayed := "Remote_Panel_DB_1".Safety_OK,
                     Safety_OK := "Remote_Panel_DB_1".Safety_Ok_Conf,
                     CNV_In_Out := "CNV_HMI".In_Out[1],
                     Cnv_Control := "Control_DB".LCnv_Sys[1].Cnv_Level[6].Cnv2,
                     SinaSpeed := "SinaSpeed_C1206_DB");
   END_IF;
   "C1207_FB_DB"(Cnv_Settings := "Settings_DB".LCnv_Sys[1].Cnv_Level[7].Cnv2,   // "Buffer_Conveyor_FB"
                 VTD_Level := "Control_DB".VTD_Sys[1].Current_Level,
                 Safety_OK_Delayed := "Remote_Panel_DB_1".Safety_OK,
                 Safety_OK := "Remote_Panel_DB_1".Safety_Ok_Conf,
                 CNV_In_Out := "CNV_HMI".In_Out[1],
                 Cnv_Control := "Control_DB".LCnv_Sys[1].Cnv_Level[7].Cnv2,
                 SinaSpeed := "SinaSpeed_C1207_DB",
                 ENO => #_w5);
   IF #_w5 THEN
       "C1208_FB_DB"(Cnv_Settings := "Settings_DB".LCnv_Sys[1].Cnv_Level[8].Cnv2,   // "Buffer_Conveyor_FB"
                     VTD_Level := "Control_DB".VTD_Sys[1].Current_Level,
                     Safety_OK_Delayed := "Remote_Panel_DB_1".Safety_OK,
                     Safety_OK := "Remote_Panel_DB_1".Safety_Ok_Conf,
                     CNV_In_Out := "CNV_HMI".In_Out[1],
                     Cnv_Control := "Control_DB".LCnv_Sys[1].Cnv_Level[8].Cnv2,
                     SinaSpeed := "SinaSpeed_C1208_DB");
   END_IF;
END_REGION

REGION Network 22: SAFETY STOPPERS Tower 1 - SYSTEM 1
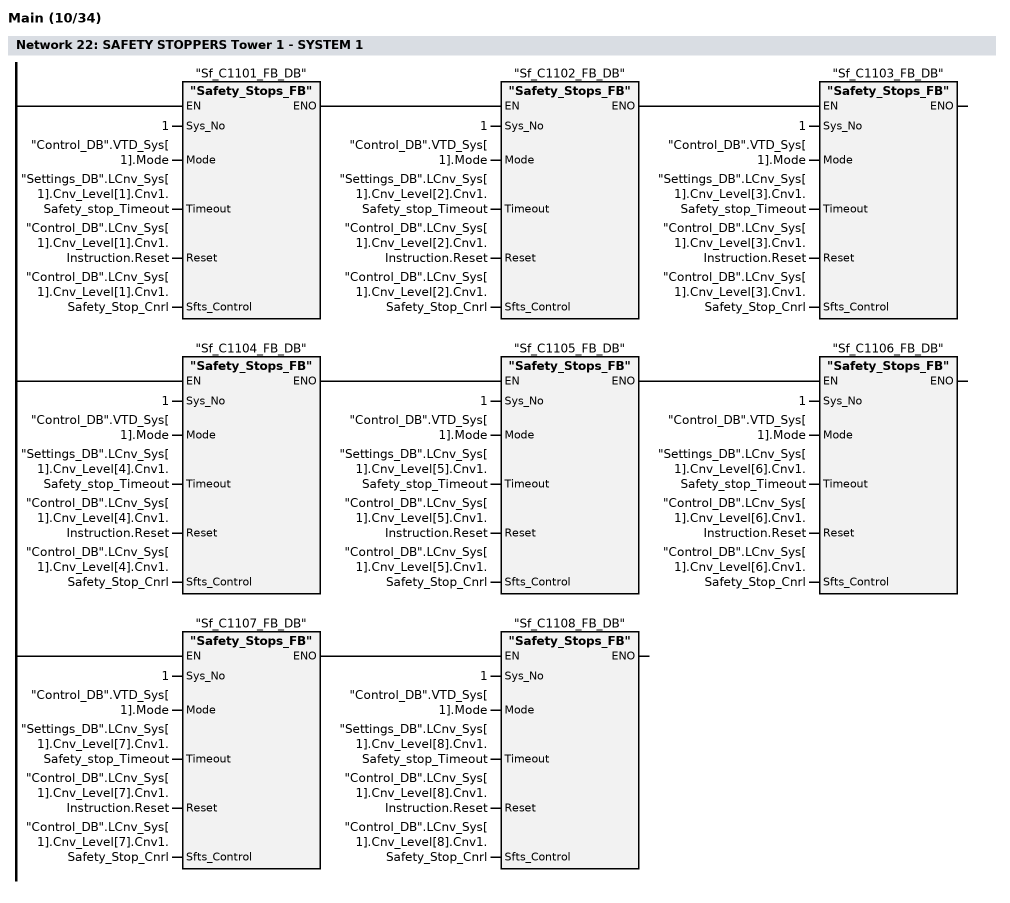
   RUNG wire#powerrail
      "Sf_C1101_FB_DB"(Sys_No := 1, Mode := "Control_DB".VTD_Sys[1].Mode, Timeout := "Settings_DB".LCnv_Sys[1].Cnv_Level[1].Cnv1.Safety_stop_Timeout, Reset := "Control_DB".LCnv_Sys[1].Cnv_Level[1].Cnv1.Instruction.Reset, Sfts_Control := "Control_DB".LCnv_Sys[1].Cnv_Level[1].Cnv1.Safety_Stop_Cnrl)
      "Sf_C1102_FB_DB"(Sys_No := 1, Mode := "Control_DB".VTD_Sys[1].Mode, Timeout := "Settings_DB".LCnv_Sys[1].Cnv_Level[2].Cnv1.Safety_stop_Timeout, Reset := "Control_DB".LCnv_Sys[1].Cnv_Level[2].Cnv1.Instruction.Reset, Sfts_Control := "Control_DB".LCnv_Sys[1].Cnv_Level[2].Cnv1.Safety_Stop_Cnrl)
      "Sf_C1103_FB_DB"(Sys_No := 1, Mode := "Control_DB".VTD_Sys[1].Mode, Timeout := "Settings_DB".LCnv_Sys[1].Cnv_Level[3].Cnv1.Safety_stop_Timeout, Reset := "Control_DB".LCnv_Sys[1].Cnv_Level[3].Cnv1.Instruction.Reset, Sfts_Control := "Control_DB".LCnv_Sys[1].Cnv_Level[3].Cnv1.Safety_Stop_Cnrl)
   END_RUNG
   RUNG wire#powerrail
      "Sf_C1104_FB_DB"(Sys_No := 1, Mode := "Control_DB".VTD_Sys[1].Mode, Timeout := "Settings_DB".LCnv_Sys[1].Cnv_Level[4].Cnv1.Safety_stop_Timeout, Reset := "Control_DB".LCnv_Sys[1].Cnv_Level[4].Cnv1.Instruction.Reset, Sfts_Control := "Control_DB".LCnv_Sys[1].Cnv_Level[4].Cnv1.Safety_Stop_Cnrl)
      "Sf_C1105_FB_DB"(Sys_No := 1, Mode := "Control_DB".VTD_Sys[1].Mode, Timeout := "Settings_DB".LCnv_Sys[1].Cnv_Level[5].Cnv1.Safety_stop_Timeout, Reset := "Control_DB".LCnv_Sys[1].Cnv_Level[5].Cnv1.Instruction.Reset, Sfts_Control := "Control_DB".LCnv_Sys[1].Cnv_Level[5].Cnv1.Safety_Stop_Cnrl)
      "Sf_C1106_FB_DB"(Sys_No := 1, Mode := "Control_DB".VTD_Sys[1].Mode, Timeout := "Settings_DB".LCnv_Sys[1].Cnv_Level[6].Cnv1.Safety_stop_Timeout, Reset := "Control_DB".LCnv_Sys[1].Cnv_Level[6].Cnv1.Instruction.Reset, Sfts_Control := "Control_DB".LCnv_Sys[1].Cnv_Level[6].Cnv1.Safety_Stop_Cnrl)
   END_RUNG
   RUNG wire#powerrail
      "Sf_C1107_FB_DB"(Sys_No := 1, Mode := "Control_DB".VTD_Sys[1].Mode, Timeout := "Settings_DB".LCnv_Sys[1].Cnv_Level[7].Cnv1.Safety_stop_Timeout, Reset := "Control_DB".LCnv_Sys[1].Cnv_Level[7].Cnv1.Instruction.Reset, Sfts_Control := "Control_DB".LCnv_Sys[1].Cnv_Level[7].Cnv1.Safety_Stop_Cnrl)
      "Sf_C1108_FB_DB"(Sys_No := 1, Mode := "Control_DB".VTD_Sys[1].Mode, Timeout := "Settings_DB".LCnv_Sys[1].Cnv_Level[8].Cnv1.Safety_stop_Timeout, Reset := "Control_DB".LCnv_Sys[1].Cnv_Level[8].Cnv1.Instruction.Reset, Sfts_Control := "Control_DB".LCnv_Sys[1].Cnv_Level[8].Cnv1.Safety_Stop_Cnrl)
   END_RUNG
   // the same network as SCL:
   "Sf_C1101_FB_DB"(Sys_No := 1,   // "Safety_Stops_FB"
                    Mode := "Control_DB".VTD_Sys[1].Mode,
                    Timeout := "Settings_DB".LCnv_Sys[1].Cnv_Level[1].Cnv1.Safety_stop_Timeout,
                    Reset := "Control_DB".LCnv_Sys[1].Cnv_Level[1].Cnv1.Instruction.Reset,
                    Sfts_Control := "Control_DB".LCnv_Sys[1].Cnv_Level[1].Cnv1.Safety_Stop_Cnrl,
                    ENO => #_w1);
   "Sf_C1102_FB_DB"(EN := #_w1,   // "Safety_Stops_FB"
                    Sys_No := 1,
                    Mode := "Control_DB".VTD_Sys[1].Mode,
                    Timeout := "Settings_DB".LCnv_Sys[1].Cnv_Level[2].Cnv1.Safety_stop_Timeout,
                    Reset := "Control_DB".LCnv_Sys[1].Cnv_Level[2].Cnv1.Instruction.Reset,
                    Sfts_Control := "Control_DB".LCnv_Sys[1].Cnv_Level[2].Cnv1.Safety_Stop_Cnrl,
                    ENO => #_w2);
   IF #_w2 THEN
       "Sf_C1103_FB_DB"(Sys_No := 1,   // "Safety_Stops_FB"
                        Mode := "Control_DB".VTD_Sys[1].Mode,
                        Timeout := "Settings_DB".LCnv_Sys[1].Cnv_Level[3].Cnv1.Safety_stop_Timeout,
                        Reset := "Control_DB".LCnv_Sys[1].Cnv_Level[3].Cnv1.Instruction.Reset,
                        Sfts_Control := "Control_DB".LCnv_Sys[1].Cnv_Level[3].Cnv1.Safety_Stop_Cnrl);
   END_IF;
   "Sf_C1104_FB_DB"(Sys_No := 1,   // "Safety_Stops_FB"
                    Mode := "Control_DB".VTD_Sys[1].Mode,
                    Timeout := "Settings_DB".LCnv_Sys[1].Cnv_Level[4].Cnv1.Safety_stop_Timeout,
                    Reset := "Control_DB".LCnv_Sys[1].Cnv_Level[4].Cnv1.Instruction.Reset,
                    Sfts_Control := "Control_DB".LCnv_Sys[1].Cnv_Level[4].Cnv1.Safety_Stop_Cnrl,
                    ENO => #_w3);
   "Sf_C1105_FB_DB"(EN := #_w3,   // "Safety_Stops_FB"
                    Sys_No := 1,
                    Mode := "Control_DB".VTD_Sys[1].Mode,
                    Timeout := "Settings_DB".LCnv_Sys[1].Cnv_Level[5].Cnv1.Safety_stop_Timeout,
                    Reset := "Control_DB".LCnv_Sys[1].Cnv_Level[5].Cnv1.Instruction.Reset,
                    Sfts_Control := "Control_DB".LCnv_Sys[1].Cnv_Level[5].Cnv1.Safety_Stop_Cnrl,
                    ENO => #_w4);
   IF #_w4 THEN
       "Sf_C1106_FB_DB"(Sys_No := 1,   // "Safety_Stops_FB"
                        Mode := "Control_DB".VTD_Sys[1].Mode,
                        Timeout := "Settings_DB".LCnv_Sys[1].Cnv_Level[6].Cnv1.Safety_stop_Timeout,
                        Reset := "Control_DB".LCnv_Sys[1].Cnv_Level[6].Cnv1.Instruction.Reset,
                        Sfts_Control := "Control_DB".LCnv_Sys[1].Cnv_Level[6].Cnv1.Safety_Stop_Cnrl);
   END_IF;
   "Sf_C1107_FB_DB"(Sys_No := 1,   // "Safety_Stops_FB"
                    Mode := "Control_DB".VTD_Sys[1].Mode,
                    Timeout := "Settings_DB".LCnv_Sys[1].Cnv_Level[7].Cnv1.Safety_stop_Timeout,
                    Reset := "Control_DB".LCnv_Sys[1].Cnv_Level[7].Cnv1.Instruction.Reset,
                    Sfts_Control := "Control_DB".LCnv_Sys[1].Cnv_Level[7].Cnv1.Safety_Stop_Cnrl,
                    ENO => #_w5);
   IF #_w5 THEN
       "Sf_C1108_FB_DB"(Sys_No := 1,   // "Safety_Stops_FB"
                        Mode := "Control_DB".VTD_Sys[1].Mode,
                        Timeout := "Settings_DB".LCnv_Sys[1].Cnv_Level[8].Cnv1.Safety_stop_Timeout,
                        Reset := "Control_DB".LCnv_Sys[1].Cnv_Level[8].Cnv1.Instruction.Reset,
                        Sfts_Control := "Control_DB".LCnv_Sys[1].Cnv_Level[8].Cnv1.Safety_Stop_Cnrl);
   END_IF;
END_REGION

REGION Network 23: SAFETY STOPPERS Tower 2 - SYSTEM 1
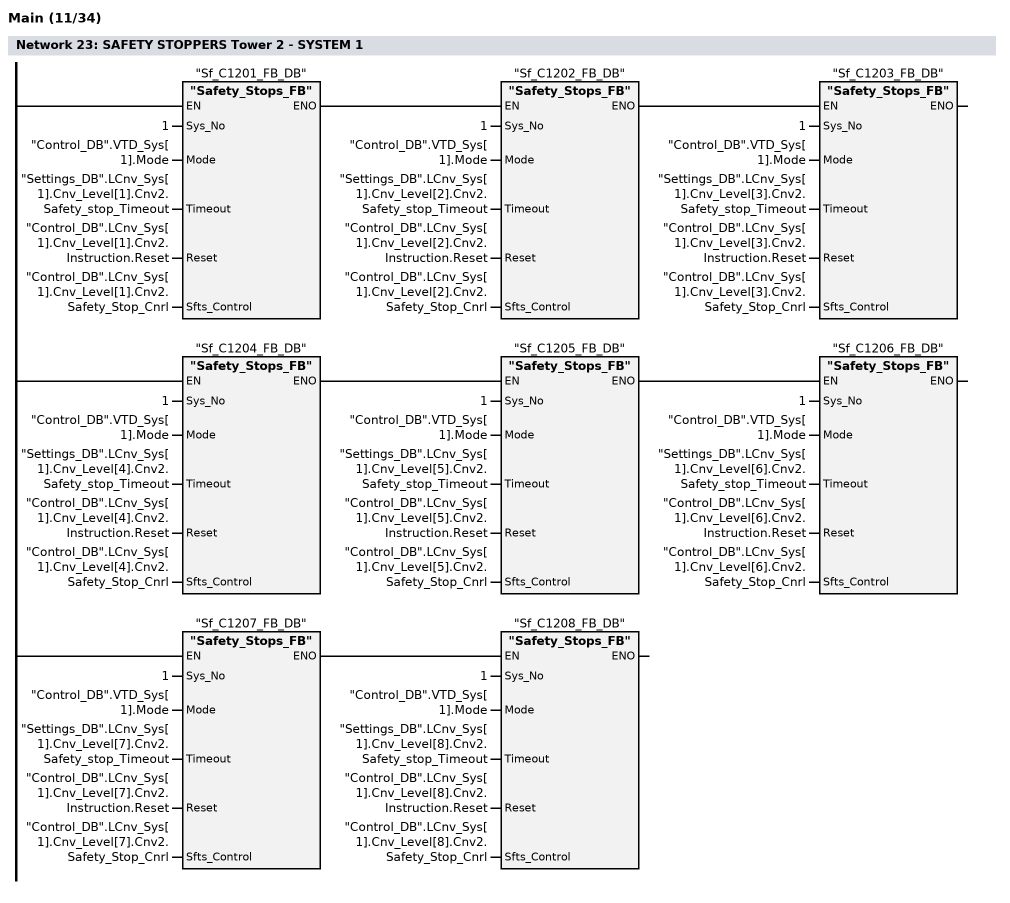
   RUNG wire#powerrail
      "Sf_C1201_FB_DB"(Sys_No := 1, Mode := "Control_DB".VTD_Sys[1].Mode, Timeout := "Settings_DB".LCnv_Sys[1].Cnv_Level[1].Cnv2.Safety_stop_Timeout, Reset := "Control_DB".LCnv_Sys[1].Cnv_Level[1].Cnv2.Instruction.Reset, Sfts_Control := "Control_DB".LCnv_Sys[1].Cnv_Level[1].Cnv2.Safety_Stop_Cnrl)
      "Sf_C1202_FB_DB"(Sys_No := 1, Mode := "Control_DB".VTD_Sys[1].Mode, Timeout := "Settings_DB".LCnv_Sys[1].Cnv_Level[2].Cnv2.Safety_stop_Timeout, Reset := "Control_DB".LCnv_Sys[1].Cnv_Level[2].Cnv2.Instruction.Reset, Sfts_Control := "Control_DB".LCnv_Sys[1].Cnv_Level[2].Cnv2.Safety_Stop_Cnrl)
      "Sf_C1203_FB_DB"(Sys_No := 1, Mode := "Control_DB".VTD_Sys[1].Mode, Timeout := "Settings_DB".LCnv_Sys[1].Cnv_Level[3].Cnv2.Safety_stop_Timeout, Reset := "Control_DB".LCnv_Sys[1].Cnv_Level[3].Cnv2.Instruction.Reset, Sfts_Control := "Control_DB".LCnv_Sys[1].Cnv_Level[3].Cnv2.Safety_Stop_Cnrl)
   END_RUNG
   RUNG wire#powerrail
      "Sf_C1204_FB_DB"(Sys_No := 1, Mode := "Control_DB".VTD_Sys[1].Mode, Timeout := "Settings_DB".LCnv_Sys[1].Cnv_Level[4].Cnv2.Safety_stop_Timeout, Reset := "Control_DB".LCnv_Sys[1].Cnv_Level[4].Cnv2.Instruction.Reset, Sfts_Control := "Control_DB".LCnv_Sys[1].Cnv_Level[4].Cnv2.Safety_Stop_Cnrl)
      "Sf_C1205_FB_DB"(Sys_No := 1, Mode := "Control_DB".VTD_Sys[1].Mode, Timeout := "Settings_DB".LCnv_Sys[1].Cnv_Level[5].Cnv2.Safety_stop_Timeout, Reset := "Control_DB".LCnv_Sys[1].Cnv_Level[5].Cnv2.Instruction.Reset, Sfts_Control := "Control_DB".LCnv_Sys[1].Cnv_Level[5].Cnv2.Safety_Stop_Cnrl)
      "Sf_C1206_FB_DB"(Sys_No := 1, Mode := "Control_DB".VTD_Sys[1].Mode, Timeout := "Settings_DB".LCnv_Sys[1].Cnv_Level[6].Cnv2.Safety_stop_Timeout, Reset := "Control_DB".LCnv_Sys[1].Cnv_Level[6].Cnv2.Instruction.Reset, Sfts_Control := "Control_DB".LCnv_Sys[1].Cnv_Level[6].Cnv2.Safety_Stop_Cnrl)
   END_RUNG
   RUNG wire#powerrail
      "Sf_C1207_FB_DB"(Sys_No := 1, Mode := "Control_DB".VTD_Sys[1].Mode, Timeout := "Settings_DB".LCnv_Sys[1].Cnv_Level[7].Cnv2.Safety_stop_Timeout, Reset := "Control_DB".LCnv_Sys[1].Cnv_Level[7].Cnv2.Instruction.Reset, Sfts_Control := "Control_DB".LCnv_Sys[1].Cnv_Level[7].Cnv2.Safety_Stop_Cnrl)
      "Sf_C1208_FB_DB"(Sys_No := 1, Mode := "Control_DB".VTD_Sys[1].Mode, Timeout := "Settings_DB".LCnv_Sys[1].Cnv_Level[8].Cnv2.Safety_stop_Timeout, Reset := "Control_DB".LCnv_Sys[1].Cnv_Level[8].Cnv2.Instruction.Reset, Sfts_Control := "Control_DB".LCnv_Sys[1].Cnv_Level[8].Cnv2.Safety_Stop_Cnrl)
   END_RUNG
   // the same network as SCL:
   "Sf_C1201_FB_DB"(Sys_No := 1,   // "Safety_Stops_FB"
                    Mode := "Control_DB".VTD_Sys[1].Mode,
                    Timeout := "Settings_DB".LCnv_Sys[1].Cnv_Level[1].Cnv2.Safety_stop_Timeout,
                    Reset := "Control_DB".LCnv_Sys[1].Cnv_Level[1].Cnv2.Instruction.Reset,
                    Sfts_Control := "Control_DB".LCnv_Sys[1].Cnv_Level[1].Cnv2.Safety_Stop_Cnrl,
                    ENO => #_w1);
   "Sf_C1202_FB_DB"(EN := #_w1,   // "Safety_Stops_FB"
                    Sys_No := 1,
                    Mode := "Control_DB".VTD_Sys[1].Mode,
                    Timeout := "Settings_DB".LCnv_Sys[1].Cnv_Level[2].Cnv2.Safety_stop_Timeout,
                    Reset := "Control_DB".LCnv_Sys[1].Cnv_Level[2].Cnv2.Instruction.Reset,
                    Sfts_Control := "Control_DB".LCnv_Sys[1].Cnv_Level[2].Cnv2.Safety_Stop_Cnrl,
                    ENO => #_w2);
   IF #_w2 THEN
       "Sf_C1203_FB_DB"(Sys_No := 1,   // "Safety_Stops_FB"
                        Mode := "Control_DB".VTD_Sys[1].Mode,
                        Timeout := "Settings_DB".LCnv_Sys[1].Cnv_Level[3].Cnv2.Safety_stop_Timeout,
                        Reset := "Control_DB".LCnv_Sys[1].Cnv_Level[3].Cnv2.Instruction.Reset,
                        Sfts_Control := "Control_DB".LCnv_Sys[1].Cnv_Level[3].Cnv2.Safety_Stop_Cnrl);
   END_IF;
   "Sf_C1204_FB_DB"(Sys_No := 1,   // "Safety_Stops_FB"
                    Mode := "Control_DB".VTD_Sys[1].Mode,
                    Timeout := "Settings_DB".LCnv_Sys[1].Cnv_Level[4].Cnv2.Safety_stop_Timeout,
                    Reset := "Control_DB".LCnv_Sys[1].Cnv_Level[4].Cnv2.Instruction.Reset,
                    Sfts_Control := "Control_DB".LCnv_Sys[1].Cnv_Level[4].Cnv2.Safety_Stop_Cnrl,
                    ENO => #_w3);
   "Sf_C1205_FB_DB"(EN := #_w3,   // "Safety_Stops_FB"
                    Sys_No := 1,
                    Mode := "Control_DB".VTD_Sys[1].Mode,
                    Timeout := "Settings_DB".LCnv_Sys[1].Cnv_Level[5].Cnv2.Safety_stop_Timeout,
                    Reset := "Control_DB".LCnv_Sys[1].Cnv_Level[5].Cnv2.Instruction.Reset,
                    Sfts_Control := "Control_DB".LCnv_Sys[1].Cnv_Level[5].Cnv2.Safety_Stop_Cnrl,
                    ENO => #_w4);
   IF #_w4 THEN
       "Sf_C1206_FB_DB"(Sys_No := 1,   // "Safety_Stops_FB"
                        Mode := "Control_DB".VTD_Sys[1].Mode,
                        Timeout := "Settings_DB".LCnv_Sys[1].Cnv_Level[6].Cnv2.Safety_stop_Timeout,
                        Reset := "Control_DB".LCnv_Sys[1].Cnv_Level[6].Cnv2.Instruction.Reset,
                        Sfts_Control := "Control_DB".LCnv_Sys[1].Cnv_Level[6].Cnv2.Safety_Stop_Cnrl);
   END_IF;
   "Sf_C1207_FB_DB"(Sys_No := 1,   // "Safety_Stops_FB"
                    Mode := "Control_DB".VTD_Sys[1].Mode,
                    Timeout := "Settings_DB".LCnv_Sys[1].Cnv_Level[7].Cnv2.Safety_stop_Timeout,
                    Reset := "Control_DB".LCnv_Sys[1].Cnv_Level[7].Cnv2.Instruction.Reset,
                    Sfts_Control := "Control_DB".LCnv_Sys[1].Cnv_Level[7].Cnv2.Safety_Stop_Cnrl,
                    ENO => #_w5);
   IF #_w5 THEN
       "Sf_C1208_FB_DB"(Sys_No := 1,   // "Safety_Stops_FB"
                        Mode := "Control_DB".VTD_Sys[1].Mode,
                        Timeout := "Settings_DB".LCnv_Sys[1].Cnv_Level[8].Cnv2.Safety_stop_Timeout,
                        Reset := "Control_DB".LCnv_Sys[1].Cnv_Level[8].Cnv2.Instruction.Reset,
                        Sfts_Control := "Control_DB".LCnv_Sys[1].Cnv_Level[8].Cnv2.Safety_Stop_Cnrl);
   END_IF;
END_REGION

REGION Network 24: SYSTEM 2
END_REGION

REGION Network 25: Level Conveyors Tower 1 - SYSTEM 2
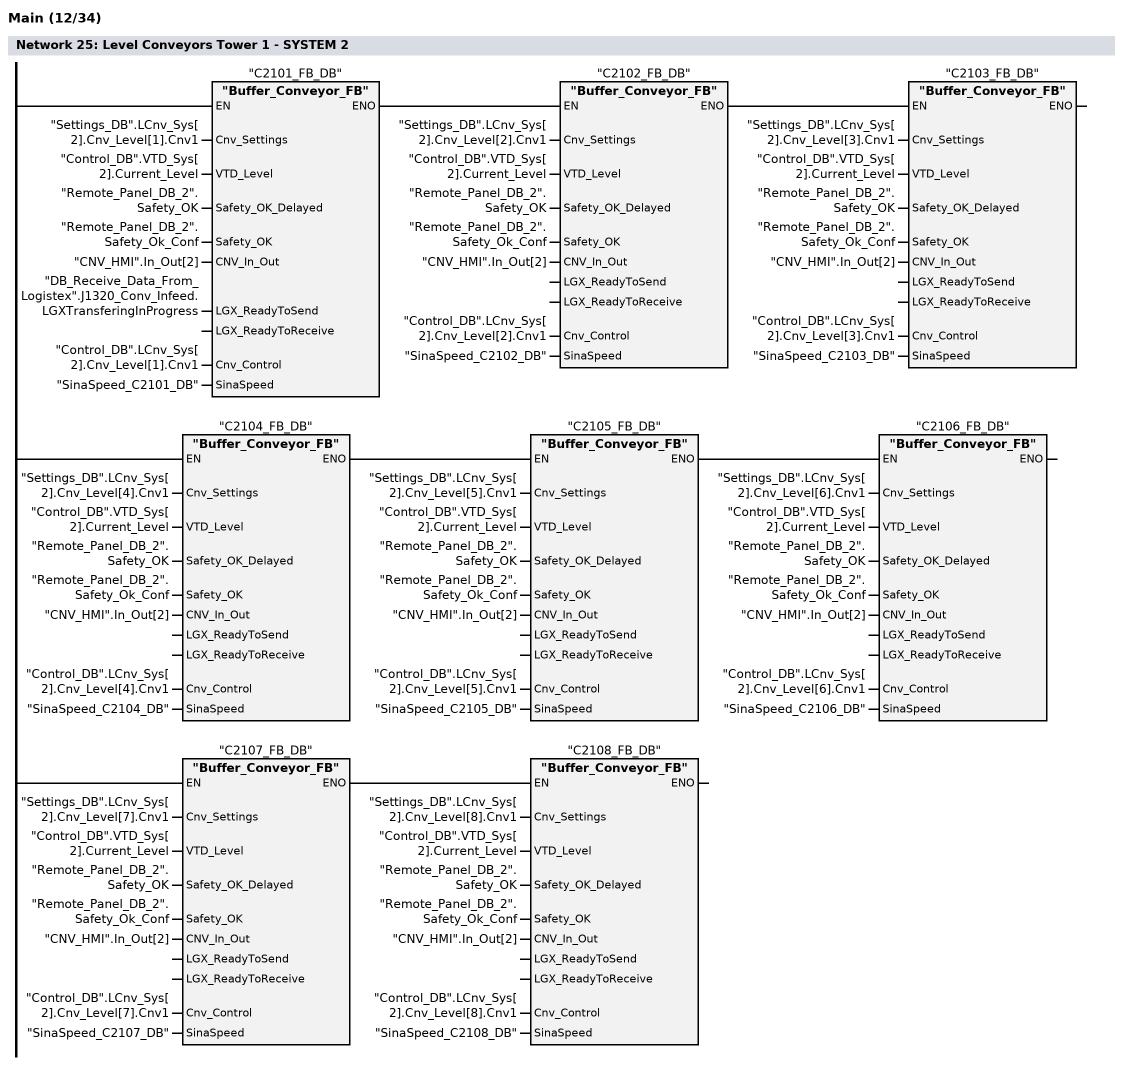
   RUNG wire#powerrail
      "C2101_FB_DB"(Cnv_Settings := "Settings_DB".LCnv_Sys[2].Cnv_Level[1].Cnv1, VTD_Level := "Control_DB".VTD_Sys[2].Current_Level, Safety_OK_Delayed := "Remote_Panel_DB_2".Safety_OK, Safety_OK := "Remote_Panel_DB_2".Safety_Ok_Conf, CNV_In_Out := "CNV_HMI".In_Out[2], LGX_ReadyToSend := "DB_Receive_Data_From_Logistex".J1320_Conv_Infeed.LGXTransferingInProgress, LGX_ReadyToReceive :=, Cnv_Control := "Control_DB".LCnv_Sys[2].Cnv_Level[1].Cnv1, SinaSpeed := "SinaSpeed_C2101_DB")
      "C2102_FB_DB"(Cnv_Settings := "Settings_DB".LCnv_Sys[2].Cnv_Level[2].Cnv1, VTD_Level := "Control_DB".VTD_Sys[2].Current_Level, Safety_OK_Delayed := "Remote_Panel_DB_2".Safety_OK, Safety_OK := "Remote_Panel_DB_2".Safety_Ok_Conf, CNV_In_Out := "CNV_HMI".In_Out[2], LGX_ReadyToSend :=, LGX_ReadyToReceive :=, Cnv_Control := "Control_DB".LCnv_Sys[2].Cnv_Level[2].Cnv1, SinaSpeed := "SinaSpeed_C2102_DB")
      "C2103_FB_DB"(Cnv_Settings := "Settings_DB".LCnv_Sys[2].Cnv_Level[3].Cnv1, VTD_Level := "Control_DB".VTD_Sys[2].Current_Level, Safety_OK_Delayed := "Remote_Panel_DB_2".Safety_OK, Safety_OK := "Remote_Panel_DB_2".Safety_Ok_Conf, CNV_In_Out := "CNV_HMI".In_Out[2], LGX_ReadyToSend :=, LGX_ReadyToReceive :=, Cnv_Control := "Control_DB".LCnv_Sys[2].Cnv_Level[3].Cnv1, SinaSpeed := "SinaSpeed_C2103_DB")
   END_RUNG
   RUNG wire#powerrail
      "C2104_FB_DB"(Cnv_Settings := "Settings_DB".LCnv_Sys[2].Cnv_Level[4].Cnv1, VTD_Level := "Control_DB".VTD_Sys[2].Current_Level, Safety_OK_Delayed := "Remote_Panel_DB_2".Safety_OK, Safety_OK := "Remote_Panel_DB_2".Safety_Ok_Conf, CNV_In_Out := "CNV_HMI".In_Out[2], LGX_ReadyToSend :=, LGX_ReadyToReceive :=, Cnv_Control := "Control_DB".LCnv_Sys[2].Cnv_Level[4].Cnv1, SinaSpeed := "SinaSpeed_C2104_DB")
      "C2105_FB_DB"(Cnv_Settings := "Settings_DB".LCnv_Sys[2].Cnv_Level[5].Cnv1, VTD_Level := "Control_DB".VTD_Sys[2].Current_Level, Safety_OK_Delayed := "Remote_Panel_DB_2".Safety_OK, Safety_OK := "Remote_Panel_DB_2".Safety_Ok_Conf, CNV_In_Out := "CNV_HMI".In_Out[2], LGX_ReadyToSend :=, LGX_ReadyToReceive :=, Cnv_Control := "Control_DB".LCnv_Sys[2].Cnv_Level[5].Cnv1, SinaSpeed := "SinaSpeed_C2105_DB")
      "C2106_FB_DB"(Cnv_Settings := "Settings_DB".LCnv_Sys[2].Cnv_Level[6].Cnv1, VTD_Level := "Control_DB".VTD_Sys[2].Current_Level, Safety_OK_Delayed := "Remote_Panel_DB_2".Safety_OK, Safety_OK := "Remote_Panel_DB_2".Safety_Ok_Conf, CNV_In_Out := "CNV_HMI".In_Out[2], LGX_ReadyToSend :=, LGX_ReadyToReceive :=, Cnv_Control := "Control_DB".LCnv_Sys[2].Cnv_Level[6].Cnv1, SinaSpeed := "SinaSpeed_C2106_DB")
   END_RUNG
   RUNG wire#powerrail
      "C2107_FB_DB"(Cnv_Settings := "Settings_DB".LCnv_Sys[2].Cnv_Level[7].Cnv1, VTD_Level := "Control_DB".VTD_Sys[2].Current_Level, Safety_OK_Delayed := "Remote_Panel_DB_2".Safety_OK, Safety_OK := "Remote_Panel_DB_2".Safety_Ok_Conf, CNV_In_Out := "CNV_HMI".In_Out[2], LGX_ReadyToSend :=, LGX_ReadyToReceive :=, Cnv_Control := "Control_DB".LCnv_Sys[2].Cnv_Level[7].Cnv1, SinaSpeed := "SinaSpeed_C2107_DB")
      "C2108_FB_DB"(Cnv_Settings := "Settings_DB".LCnv_Sys[2].Cnv_Level[8].Cnv1, VTD_Level := "Control_DB".VTD_Sys[2].Current_Level, Safety_OK_Delayed := "Remote_Panel_DB_2".Safety_OK, Safety_OK := "Remote_Panel_DB_2".Safety_Ok_Conf, CNV_In_Out := "CNV_HMI".In_Out[2], LGX_ReadyToSend :=, LGX_ReadyToReceive :=, Cnv_Control := "Control_DB".LCnv_Sys[2].Cnv_Level[8].Cnv1, SinaSpeed := "SinaSpeed_C2108_DB")
   END_RUNG
   // the same network as SCL:
   "C2101_FB_DB"(Cnv_Settings := "Settings_DB".LCnv_Sys[2].Cnv_Level[1].Cnv1,   // "Buffer_Conveyor_FB"
                 VTD_Level := "Control_DB".VTD_Sys[2].Current_Level,
                 Safety_OK_Delayed := "Remote_Panel_DB_2".Safety_OK,
                 Safety_OK := "Remote_Panel_DB_2".Safety_Ok_Conf,
                 CNV_In_Out := "CNV_HMI".In_Out[2],
                 LGX_ReadyToSend := "DB_Receive_Data_From_Logistex".J1320_Conv_Infeed.LGXTransferingInProgress,
                 Cnv_Control := "Control_DB".LCnv_Sys[2].Cnv_Level[1].Cnv1,
                 SinaSpeed := "SinaSpeed_C2101_DB",
                 ENO => #_w1);
   "C2102_FB_DB"(EN := #_w1,   // "Buffer_Conveyor_FB"
                 Cnv_Settings := "Settings_DB".LCnv_Sys[2].Cnv_Level[2].Cnv1,
                 VTD_Level := "Control_DB".VTD_Sys[2].Current_Level,
                 Safety_OK_Delayed := "Remote_Panel_DB_2".Safety_OK,
                 Safety_OK := "Remote_Panel_DB_2".Safety_Ok_Conf,
                 CNV_In_Out := "CNV_HMI".In_Out[2],
                 Cnv_Control := "Control_DB".LCnv_Sys[2].Cnv_Level[2].Cnv1,
                 SinaSpeed := "SinaSpeed_C2102_DB",
                 ENO => #_w2);
   IF #_w2 THEN
       "C2103_FB_DB"(Cnv_Settings := "Settings_DB".LCnv_Sys[2].Cnv_Level[3].Cnv1,   // "Buffer_Conveyor_FB"
                     VTD_Level := "Control_DB".VTD_Sys[2].Current_Level,
                     Safety_OK_Delayed := "Remote_Panel_DB_2".Safety_OK,
                     Safety_OK := "Remote_Panel_DB_2".Safety_Ok_Conf,
                     CNV_In_Out := "CNV_HMI".In_Out[2],
                     Cnv_Control := "Control_DB".LCnv_Sys[2].Cnv_Level[3].Cnv1,
                     SinaSpeed := "SinaSpeed_C2103_DB");
   END_IF;
   "C2104_FB_DB"(Cnv_Settings := "Settings_DB".LCnv_Sys[2].Cnv_Level[4].Cnv1,   // "Buffer_Conveyor_FB"
                 VTD_Level := "Control_DB".VTD_Sys[2].Current_Level,
                 Safety_OK_Delayed := "Remote_Panel_DB_2".Safety_OK,
                 Safety_OK := "Remote_Panel_DB_2".Safety_Ok_Conf,
                 CNV_In_Out := "CNV_HMI".In_Out[2],
                 Cnv_Control := "Control_DB".LCnv_Sys[2].Cnv_Level[4].Cnv1,
                 SinaSpeed := "SinaSpeed_C2104_DB",
                 ENO => #_w3);
   "C2105_FB_DB"(EN := #_w3,   // "Buffer_Conveyor_FB"
                 Cnv_Settings := "Settings_DB".LCnv_Sys[2].Cnv_Level[5].Cnv1,
                 VTD_Level := "Control_DB".VTD_Sys[2].Current_Level,
                 Safety_OK_Delayed := "Remote_Panel_DB_2".Safety_OK,
                 Safety_OK := "Remote_Panel_DB_2".Safety_Ok_Conf,
                 CNV_In_Out := "CNV_HMI".In_Out[2],
                 Cnv_Control := "Control_DB".LCnv_Sys[2].Cnv_Level[5].Cnv1,
                 SinaSpeed := "SinaSpeed_C2105_DB",
                 ENO => #_w4);
   IF #_w4 THEN
       "C2106_FB_DB"(Cnv_Settings := "Settings_DB".LCnv_Sys[2].Cnv_Level[6].Cnv1,   // "Buffer_Conveyor_FB"
                     VTD_Level := "Control_DB".VTD_Sys[2].Current_Level,
                     Safety_OK_Delayed := "Remote_Panel_DB_2".Safety_OK,
                     Safety_OK := "Remote_Panel_DB_2".Safety_Ok_Conf,
                     CNV_In_Out := "CNV_HMI".In_Out[2],
                     Cnv_Control := "Control_DB".LCnv_Sys[2].Cnv_Level[6].Cnv1,
                     SinaSpeed := "SinaSpeed_C2106_DB");
   END_IF;
   "C2107_FB_DB"(Cnv_Settings := "Settings_DB".LCnv_Sys[2].Cnv_Level[7].Cnv1,   // "Buffer_Conveyor_FB"
                 VTD_Level := "Control_DB".VTD_Sys[2].Current_Level,
                 Safety_OK_Delayed := "Remote_Panel_DB_2".Safety_OK,
                 Safety_OK := "Remote_Panel_DB_2".Safety_Ok_Conf,
                 CNV_In_Out := "CNV_HMI".In_Out[2],
                 Cnv_Control := "Control_DB".LCnv_Sys[2].Cnv_Level[7].Cnv1,
                 SinaSpeed := "SinaSpeed_C2107_DB",
                 ENO => #_w5);
   IF #_w5 THEN
       "C2108_FB_DB"(Cnv_Settings := "Settings_DB".LCnv_Sys[2].Cnv_Level[8].Cnv1,   // "Buffer_Conveyor_FB"
                     VTD_Level := "Control_DB".VTD_Sys[2].Current_Level,
                     Safety_OK_Delayed := "Remote_Panel_DB_2".Safety_OK,
                     Safety_OK := "Remote_Panel_DB_2".Safety_Ok_Conf,
                     CNV_In_Out := "CNV_HMI".In_Out[2],
                     Cnv_Control := "Control_DB".LCnv_Sys[2].Cnv_Level[8].Cnv1,
                     SinaSpeed := "SinaSpeed_C2108_DB");
   END_IF;
END_REGION

REGION Network 26: Level Conveyors Tower 2 - SYSTEM 2
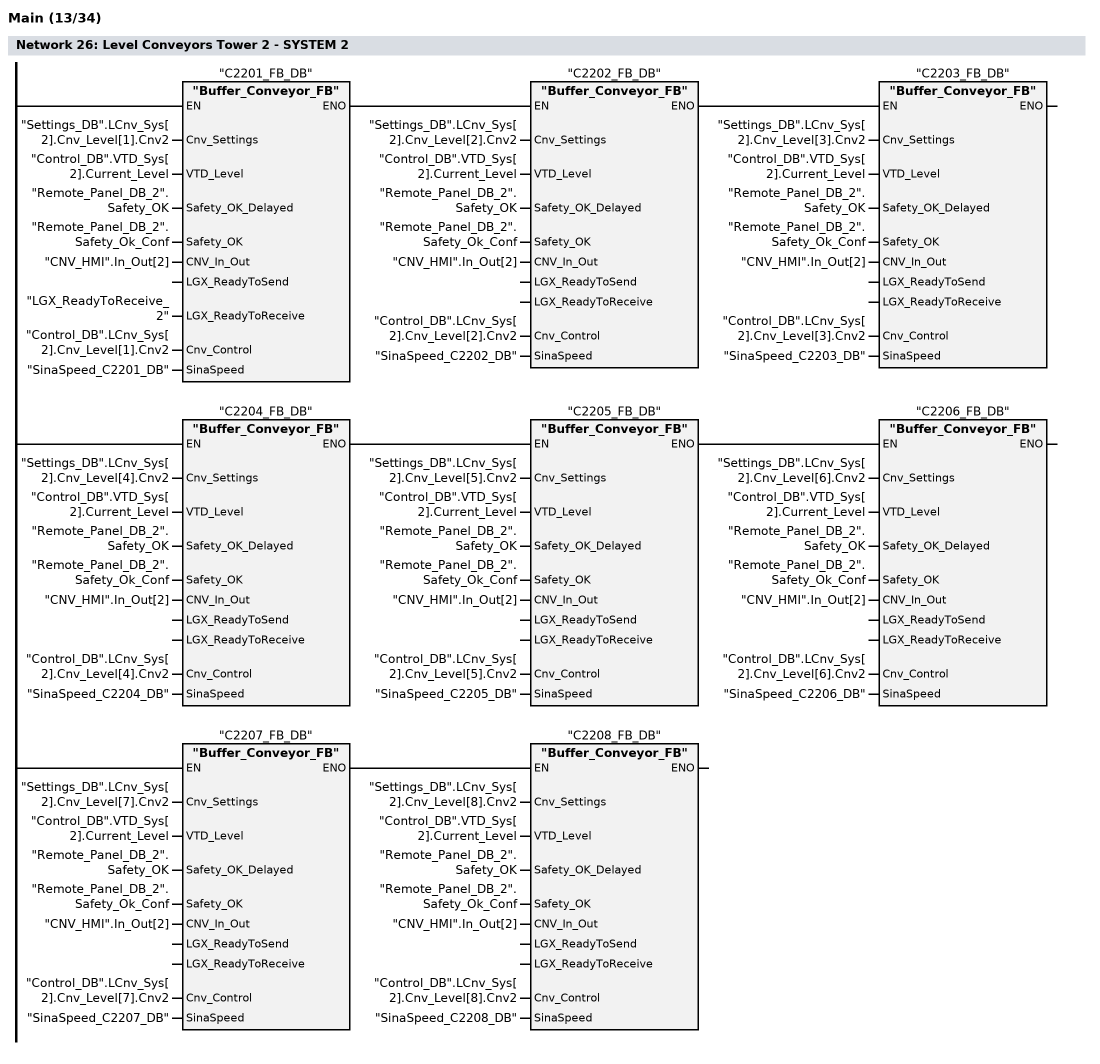
   RUNG wire#powerrail
      "C2201_FB_DB"(Cnv_Settings := "Settings_DB".LCnv_Sys[2].Cnv_Level[1].Cnv2, VTD_Level := "Control_DB".VTD_Sys[2].Current_Level, Safety_OK_Delayed := "Remote_Panel_DB_2".Safety_OK, Safety_OK := "Remote_Panel_DB_2".Safety_Ok_Conf, CNV_In_Out := "CNV_HMI".In_Out[2], LGX_ReadyToSend :=, LGX_ReadyToReceive := "LGX_ReadyToReceive_2", Cnv_Control := "Control_DB".LCnv_Sys[2].Cnv_Level[1].Cnv2, SinaSpeed := "SinaSpeed_C2201_DB")
      "C2202_FB_DB"(Cnv_Settings := "Settings_DB".LCnv_Sys[2].Cnv_Level[2].Cnv2, VTD_Level := "Control_DB".VTD_Sys[2].Current_Level, Safety_OK_Delayed := "Remote_Panel_DB_2".Safety_OK, Safety_OK := "Remote_Panel_DB_2".Safety_Ok_Conf, CNV_In_Out := "CNV_HMI".In_Out[2], LGX_ReadyToSend :=, LGX_ReadyToReceive :=, Cnv_Control := "Control_DB".LCnv_Sys[2].Cnv_Level[2].Cnv2, SinaSpeed := "SinaSpeed_C2202_DB")
      "C2203_FB_DB"(Cnv_Settings := "Settings_DB".LCnv_Sys[2].Cnv_Level[3].Cnv2, VTD_Level := "Control_DB".VTD_Sys[2].Current_Level, Safety_OK_Delayed := "Remote_Panel_DB_2".Safety_OK, Safety_OK := "Remote_Panel_DB_2".Safety_Ok_Conf, CNV_In_Out := "CNV_HMI".In_Out[2], LGX_ReadyToSend :=, LGX_ReadyToReceive :=, Cnv_Control := "Control_DB".LCnv_Sys[2].Cnv_Level[3].Cnv2, SinaSpeed := "SinaSpeed_C2203_DB")
   END_RUNG
   RUNG wire#powerrail
      "C2204_FB_DB"(Cnv_Settings := "Settings_DB".LCnv_Sys[2].Cnv_Level[4].Cnv2, VTD_Level := "Control_DB".VTD_Sys[2].Current_Level, Safety_OK_Delayed := "Remote_Panel_DB_2".Safety_OK, Safety_OK := "Remote_Panel_DB_2".Safety_Ok_Conf, CNV_In_Out := "CNV_HMI".In_Out[2], LGX_ReadyToSend :=, LGX_ReadyToReceive :=, Cnv_Control := "Control_DB".LCnv_Sys[2].Cnv_Level[4].Cnv2, SinaSpeed := "SinaSpeed_C2204_DB")
      "C2205_FB_DB"(Cnv_Settings := "Settings_DB".LCnv_Sys[2].Cnv_Level[5].Cnv2, VTD_Level := "Control_DB".VTD_Sys[2].Current_Level, Safety_OK_Delayed := "Remote_Panel_DB_2".Safety_OK, Safety_OK := "Remote_Panel_DB_2".Safety_Ok_Conf, CNV_In_Out := "CNV_HMI".In_Out[2], LGX_ReadyToSend :=, LGX_ReadyToReceive :=, Cnv_Control := "Control_DB".LCnv_Sys[2].Cnv_Level[5].Cnv2, SinaSpeed := "SinaSpeed_C2205_DB")
      "C2206_FB_DB"(Cnv_Settings := "Settings_DB".LCnv_Sys[2].Cnv_Level[6].Cnv2, VTD_Level := "Control_DB".VTD_Sys[2].Current_Level, Safety_OK_Delayed := "Remote_Panel_DB_2".Safety_OK, Safety_OK := "Remote_Panel_DB_2".Safety_Ok_Conf, CNV_In_Out := "CNV_HMI".In_Out[2], LGX_ReadyToSend :=, LGX_ReadyToReceive :=, Cnv_Control := "Control_DB".LCnv_Sys[2].Cnv_Level[6].Cnv2, SinaSpeed := "SinaSpeed_C2206_DB")
   END_RUNG
   RUNG wire#powerrail
      "C2207_FB_DB"(Cnv_Settings := "Settings_DB".LCnv_Sys[2].Cnv_Level[7].Cnv2, VTD_Level := "Control_DB".VTD_Sys[2].Current_Level, Safety_OK_Delayed := "Remote_Panel_DB_2".Safety_OK, Safety_OK := "Remote_Panel_DB_2".Safety_Ok_Conf, CNV_In_Out := "CNV_HMI".In_Out[2], LGX_ReadyToSend :=, LGX_ReadyToReceive :=, Cnv_Control := "Control_DB".LCnv_Sys[2].Cnv_Level[7].Cnv2, SinaSpeed := "SinaSpeed_C2207_DB")
      "C2208_FB_DB"(Cnv_Settings := "Settings_DB".LCnv_Sys[2].Cnv_Level[8].Cnv2, VTD_Level := "Control_DB".VTD_Sys[2].Current_Level, Safety_OK_Delayed := "Remote_Panel_DB_2".Safety_OK, Safety_OK := "Remote_Panel_DB_2".Safety_Ok_Conf, CNV_In_Out := "CNV_HMI".In_Out[2], LGX_ReadyToSend :=, LGX_ReadyToReceive :=, Cnv_Control := "Control_DB".LCnv_Sys[2].Cnv_Level[8].Cnv2, SinaSpeed := "SinaSpeed_C2208_DB")
   END_RUNG
   // the same network as SCL:
   "C2201_FB_DB"(Cnv_Settings := "Settings_DB".LCnv_Sys[2].Cnv_Level[1].Cnv2,   // "Buffer_Conveyor_FB"
                 VTD_Level := "Control_DB".VTD_Sys[2].Current_Level,
                 Safety_OK_Delayed := "Remote_Panel_DB_2".Safety_OK,
                 Safety_OK := "Remote_Panel_DB_2".Safety_Ok_Conf,
                 CNV_In_Out := "CNV_HMI".In_Out[2],
                 LGX_ReadyToReceive := "LGX_ReadyToReceive_2",
                 Cnv_Control := "Control_DB".LCnv_Sys[2].Cnv_Level[1].Cnv2,
                 SinaSpeed := "SinaSpeed_C2201_DB",
                 ENO => #_w1);
   "C2202_FB_DB"(EN := #_w1,   // "Buffer_Conveyor_FB"
                 Cnv_Settings := "Settings_DB".LCnv_Sys[2].Cnv_Level[2].Cnv2,
                 VTD_Level := "Control_DB".VTD_Sys[2].Current_Level,
                 Safety_OK_Delayed := "Remote_Panel_DB_2".Safety_OK,
                 Safety_OK := "Remote_Panel_DB_2".Safety_Ok_Conf,
                 CNV_In_Out := "CNV_HMI".In_Out[2],
                 Cnv_Control := "Control_DB".LCnv_Sys[2].Cnv_Level[2].Cnv2,
                 SinaSpeed := "SinaSpeed_C2202_DB",
                 ENO => #_w2);
   IF #_w2 THEN
       "C2203_FB_DB"(Cnv_Settings := "Settings_DB".LCnv_Sys[2].Cnv_Level[3].Cnv2,   // "Buffer_Conveyor_FB"
                     VTD_Level := "Control_DB".VTD_Sys[2].Current_Level,
                     Safety_OK_Delayed := "Remote_Panel_DB_2".Safety_OK,
                     Safety_OK := "Remote_Panel_DB_2".Safety_Ok_Conf,
                     CNV_In_Out := "CNV_HMI".In_Out[2],
                     Cnv_Control := "Control_DB".LCnv_Sys[2].Cnv_Level[3].Cnv2,
                     SinaSpeed := "SinaSpeed_C2203_DB");
   END_IF;
   "C2204_FB_DB"(Cnv_Settings := "Settings_DB".LCnv_Sys[2].Cnv_Level[4].Cnv2,   // "Buffer_Conveyor_FB"
                 VTD_Level := "Control_DB".VTD_Sys[2].Current_Level,
                 Safety_OK_Delayed := "Remote_Panel_DB_2".Safety_OK,
                 Safety_OK := "Remote_Panel_DB_2".Safety_Ok_Conf,
                 CNV_In_Out := "CNV_HMI".In_Out[2],
                 Cnv_Control := "Control_DB".LCnv_Sys[2].Cnv_Level[4].Cnv2,
                 SinaSpeed := "SinaSpeed_C2204_DB",
                 ENO => #_w3);
   "C2205_FB_DB"(EN := #_w3,   // "Buffer_Conveyor_FB"
                 Cnv_Settings := "Settings_DB".LCnv_Sys[2].Cnv_Level[5].Cnv2,
                 VTD_Level := "Control_DB".VTD_Sys[2].Current_Level,
                 Safety_OK_Delayed := "Remote_Panel_DB_2".Safety_OK,
                 Safety_OK := "Remote_Panel_DB_2".Safety_Ok_Conf,
                 CNV_In_Out := "CNV_HMI".In_Out[2],
                 Cnv_Control := "Control_DB".LCnv_Sys[2].Cnv_Level[5].Cnv2,
                 SinaSpeed := "SinaSpeed_C2205_DB",
                 ENO => #_w4);
   IF #_w4 THEN
       "C2206_FB_DB"(Cnv_Settings := "Settings_DB".LCnv_Sys[2].Cnv_Level[6].Cnv2,   // "Buffer_Conveyor_FB"
                     VTD_Level := "Control_DB".VTD_Sys[2].Current_Level,
                     Safety_OK_Delayed := "Remote_Panel_DB_2".Safety_OK,
                     Safety_OK := "Remote_Panel_DB_2".Safety_Ok_Conf,
                     CNV_In_Out := "CNV_HMI".In_Out[2],
                     Cnv_Control := "Control_DB".LCnv_Sys[2].Cnv_Level[6].Cnv2,
                     SinaSpeed := "SinaSpeed_C2206_DB");
   END_IF;
   "C2207_FB_DB"(Cnv_Settings := "Settings_DB".LCnv_Sys[2].Cnv_Level[7].Cnv2,   // "Buffer_Conveyor_FB"
                 VTD_Level := "Control_DB".VTD_Sys[2].Current_Level,
                 Safety_OK_Delayed := "Remote_Panel_DB_2".Safety_OK,
                 Safety_OK := "Remote_Panel_DB_2".Safety_Ok_Conf,
                 CNV_In_Out := "CNV_HMI".In_Out[2],
                 Cnv_Control := "Control_DB".LCnv_Sys[2].Cnv_Level[7].Cnv2,
                 SinaSpeed := "SinaSpeed_C2207_DB",
                 ENO => #_w5);
   IF #_w5 THEN
       "C2208_FB_DB"(Cnv_Settings := "Settings_DB".LCnv_Sys[2].Cnv_Level[8].Cnv2,   // "Buffer_Conveyor_FB"
                     VTD_Level := "Control_DB".VTD_Sys[2].Current_Level,
                     Safety_OK_Delayed := "Remote_Panel_DB_2".Safety_OK,
                     Safety_OK := "Remote_Panel_DB_2".Safety_Ok_Conf,
                     CNV_In_Out := "CNV_HMI".In_Out[2],
                     Cnv_Control := "Control_DB".LCnv_Sys[2].Cnv_Level[8].Cnv2,
                     SinaSpeed := "SinaSpeed_C2208_DB");
   END_IF;
END_REGION

REGION Network 27: SAFETY STOPPERS Tower 1 - SYSTEM 2
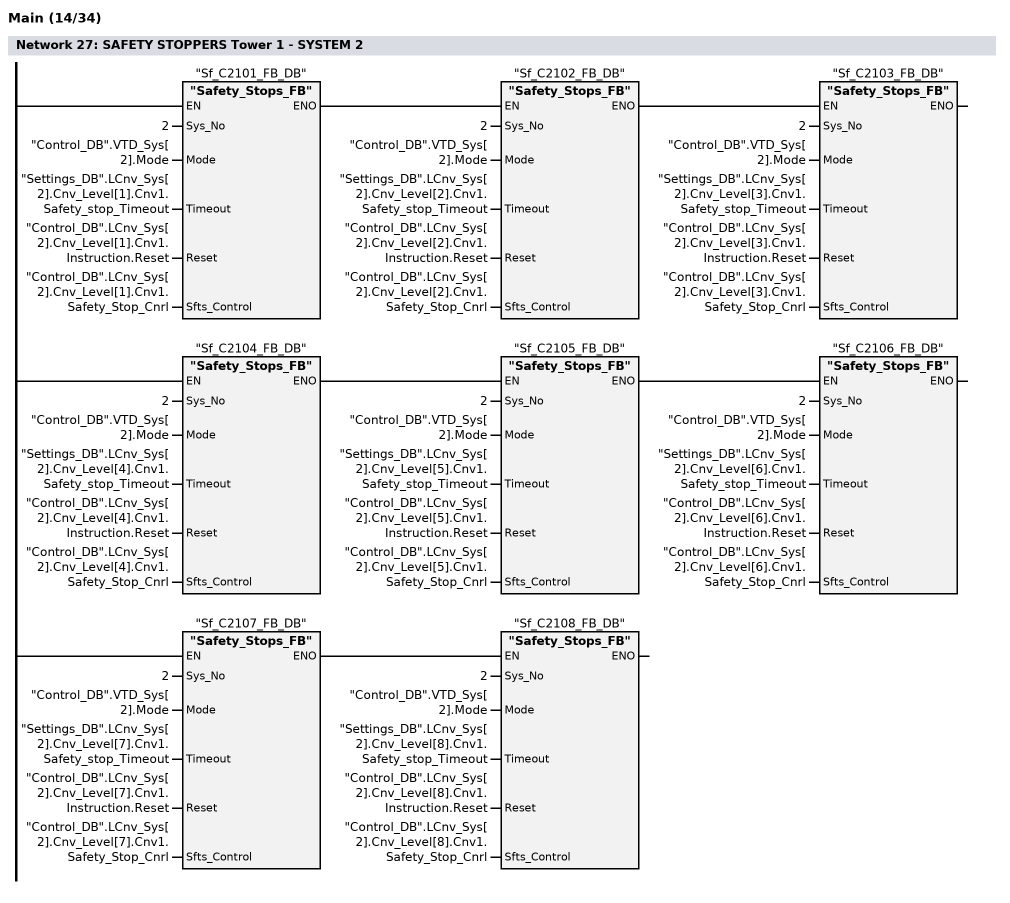
   RUNG wire#powerrail
      "Sf_C2101_FB_DB"(Sys_No := 2, Mode := "Control_DB".VTD_Sys[2].Mode, Timeout := "Settings_DB".LCnv_Sys[2].Cnv_Level[1].Cnv1.Safety_stop_Timeout, Reset := "Control_DB".LCnv_Sys[2].Cnv_Level[1].Cnv1.Instruction.Reset, Sfts_Control := "Control_DB".LCnv_Sys[2].Cnv_Level[1].Cnv1.Safety_Stop_Cnrl)
      "Sf_C2102_FB_DB"(Sys_No := 2, Mode := "Control_DB".VTD_Sys[2].Mode, Timeout := "Settings_DB".LCnv_Sys[2].Cnv_Level[2].Cnv1.Safety_stop_Timeout, Reset := "Control_DB".LCnv_Sys[2].Cnv_Level[2].Cnv1.Instruction.Reset, Sfts_Control := "Control_DB".LCnv_Sys[2].Cnv_Level[2].Cnv1.Safety_Stop_Cnrl)
      "Sf_C2103_FB_DB"(Sys_No := 2, Mode := "Control_DB".VTD_Sys[2].Mode, Timeout := "Settings_DB".LCnv_Sys[2].Cnv_Level[3].Cnv1.Safety_stop_Timeout, Reset := "Control_DB".LCnv_Sys[2].Cnv_Level[3].Cnv1.Instruction.Reset, Sfts_Control := "Control_DB".LCnv_Sys[2].Cnv_Level[3].Cnv1.Safety_Stop_Cnrl)
   END_RUNG
   RUNG wire#powerrail
      "Sf_C2104_FB_DB"(Sys_No := 2, Mode := "Control_DB".VTD_Sys[2].Mode, Timeout := "Settings_DB".LCnv_Sys[2].Cnv_Level[4].Cnv1.Safety_stop_Timeout, Reset := "Control_DB".LCnv_Sys[2].Cnv_Level[4].Cnv1.Instruction.Reset, Sfts_Control := "Control_DB".LCnv_Sys[2].Cnv_Level[4].Cnv1.Safety_Stop_Cnrl)
      "Sf_C2105_FB_DB"(Sys_No := 2, Mode := "Control_DB".VTD_Sys[2].Mode, Timeout := "Settings_DB".LCnv_Sys[2].Cnv_Level[5].Cnv1.Safety_stop_Timeout, Reset := "Control_DB".LCnv_Sys[2].Cnv_Level[5].Cnv1.Instruction.Reset, Sfts_Control := "Control_DB".LCnv_Sys[2].Cnv_Level[5].Cnv1.Safety_Stop_Cnrl)
      "Sf_C2106_FB_DB"(Sys_No := 2, Mode := "Control_DB".VTD_Sys[2].Mode, Timeout := "Settings_DB".LCnv_Sys[2].Cnv_Level[6].Cnv1.Safety_stop_Timeout, Reset := "Control_DB".LCnv_Sys[2].Cnv_Level[6].Cnv1.Instruction.Reset, Sfts_Control := "Control_DB".LCnv_Sys[2].Cnv_Level[6].Cnv1.Safety_Stop_Cnrl)
   END_RUNG
   RUNG wire#powerrail
      "Sf_C2107_FB_DB"(Sys_No := 2, Mode := "Control_DB".VTD_Sys[2].Mode, Timeout := "Settings_DB".LCnv_Sys[2].Cnv_Level[7].Cnv1.Safety_stop_Timeout, Reset := "Control_DB".LCnv_Sys[2].Cnv_Level[7].Cnv1.Instruction.Reset, Sfts_Control := "Control_DB".LCnv_Sys[2].Cnv_Level[7].Cnv1.Safety_Stop_Cnrl)
      "Sf_C2108_FB_DB"(Sys_No := 2, Mode := "Control_DB".VTD_Sys[2].Mode, Timeout := "Settings_DB".LCnv_Sys[2].Cnv_Level[8].Cnv1.Safety_stop_Timeout, Reset := "Control_DB".LCnv_Sys[2].Cnv_Level[8].Cnv1.Instruction.Reset, Sfts_Control := "Control_DB".LCnv_Sys[2].Cnv_Level[8].Cnv1.Safety_Stop_Cnrl)
   END_RUNG
   // the same network as SCL:
   "Sf_C2101_FB_DB"(Sys_No := 2,   // "Safety_Stops_FB"
                    Mode := "Control_DB".VTD_Sys[2].Mode,
                    Timeout := "Settings_DB".LCnv_Sys[2].Cnv_Level[1].Cnv1.Safety_stop_Timeout,
                    Reset := "Control_DB".LCnv_Sys[2].Cnv_Level[1].Cnv1.Instruction.Reset,
                    Sfts_Control := "Control_DB".LCnv_Sys[2].Cnv_Level[1].Cnv1.Safety_Stop_Cnrl,
                    ENO => #_w1);
   "Sf_C2102_FB_DB"(EN := #_w1,   // "Safety_Stops_FB"
                    Sys_No := 2,
                    Mode := "Control_DB".VTD_Sys[2].Mode,
                    Timeout := "Settings_DB".LCnv_Sys[2].Cnv_Level[2].Cnv1.Safety_stop_Timeout,
                    Reset := "Control_DB".LCnv_Sys[2].Cnv_Level[2].Cnv1.Instruction.Reset,
                    Sfts_Control := "Control_DB".LCnv_Sys[2].Cnv_Level[2].Cnv1.Safety_Stop_Cnrl,
                    ENO => #_w2);
   IF #_w2 THEN
       "Sf_C2103_FB_DB"(Sys_No := 2,   // "Safety_Stops_FB"
                        Mode := "Control_DB".VTD_Sys[2].Mode,
                        Timeout := "Settings_DB".LCnv_Sys[2].Cnv_Level[3].Cnv1.Safety_stop_Timeout,
                        Reset := "Control_DB".LCnv_Sys[2].Cnv_Level[3].Cnv1.Instruction.Reset,
                        Sfts_Control := "Control_DB".LCnv_Sys[2].Cnv_Level[3].Cnv1.Safety_Stop_Cnrl);
   END_IF;
   "Sf_C2104_FB_DB"(Sys_No := 2,   // "Safety_Stops_FB"
                    Mode := "Control_DB".VTD_Sys[2].Mode,
                    Timeout := "Settings_DB".LCnv_Sys[2].Cnv_Level[4].Cnv1.Safety_stop_Timeout,
                    Reset := "Control_DB".LCnv_Sys[2].Cnv_Level[4].Cnv1.Instruction.Reset,
                    Sfts_Control := "Control_DB".LCnv_Sys[2].Cnv_Level[4].Cnv1.Safety_Stop_Cnrl,
                    ENO => #_w3);
   "Sf_C2105_FB_DB"(EN := #_w3,   // "Safety_Stops_FB"
                    Sys_No := 2,
                    Mode := "Control_DB".VTD_Sys[2].Mode,
                    Timeout := "Settings_DB".LCnv_Sys[2].Cnv_Level[5].Cnv1.Safety_stop_Timeout,
                    Reset := "Control_DB".LCnv_Sys[2].Cnv_Level[5].Cnv1.Instruction.Reset,
                    Sfts_Control := "Control_DB".LCnv_Sys[2].Cnv_Level[5].Cnv1.Safety_Stop_Cnrl,
                    ENO => #_w4);
   IF #_w4 THEN
       "Sf_C2106_FB_DB"(Sys_No := 2,   // "Safety_Stops_FB"
                        Mode := "Control_DB".VTD_Sys[2].Mode,
                        Timeout := "Settings_DB".LCnv_Sys[2].Cnv_Level[6].Cnv1.Safety_stop_Timeout,
                        Reset := "Control_DB".LCnv_Sys[2].Cnv_Level[6].Cnv1.Instruction.Reset,
                        Sfts_Control := "Control_DB".LCnv_Sys[2].Cnv_Level[6].Cnv1.Safety_Stop_Cnrl);
   END_IF;
   "Sf_C2107_FB_DB"(Sys_No := 2,   // "Safety_Stops_FB"
                    Mode := "Control_DB".VTD_Sys[2].Mode,
                    Timeout := "Settings_DB".LCnv_Sys[2].Cnv_Level[7].Cnv1.Safety_stop_Timeout,
                    Reset := "Control_DB".LCnv_Sys[2].Cnv_Level[7].Cnv1.Instruction.Reset,
                    Sfts_Control := "Control_DB".LCnv_Sys[2].Cnv_Level[7].Cnv1.Safety_Stop_Cnrl,
                    ENO => #_w5);
   IF #_w5 THEN
       "Sf_C2108_FB_DB"(Sys_No := 2,   // "Safety_Stops_FB"
                        Mode := "Control_DB".VTD_Sys[2].Mode,
                        Timeout := "Settings_DB".LCnv_Sys[2].Cnv_Level[8].Cnv1.Safety_stop_Timeout,
                        Reset := "Control_DB".LCnv_Sys[2].Cnv_Level[8].Cnv1.Instruction.Reset,
                        Sfts_Control := "Control_DB".LCnv_Sys[2].Cnv_Level[8].Cnv1.Safety_Stop_Cnrl);
   END_IF;
END_REGION

REGION Network 28: SAFETY STOPPERS Tower 2 - SYSTEM 2
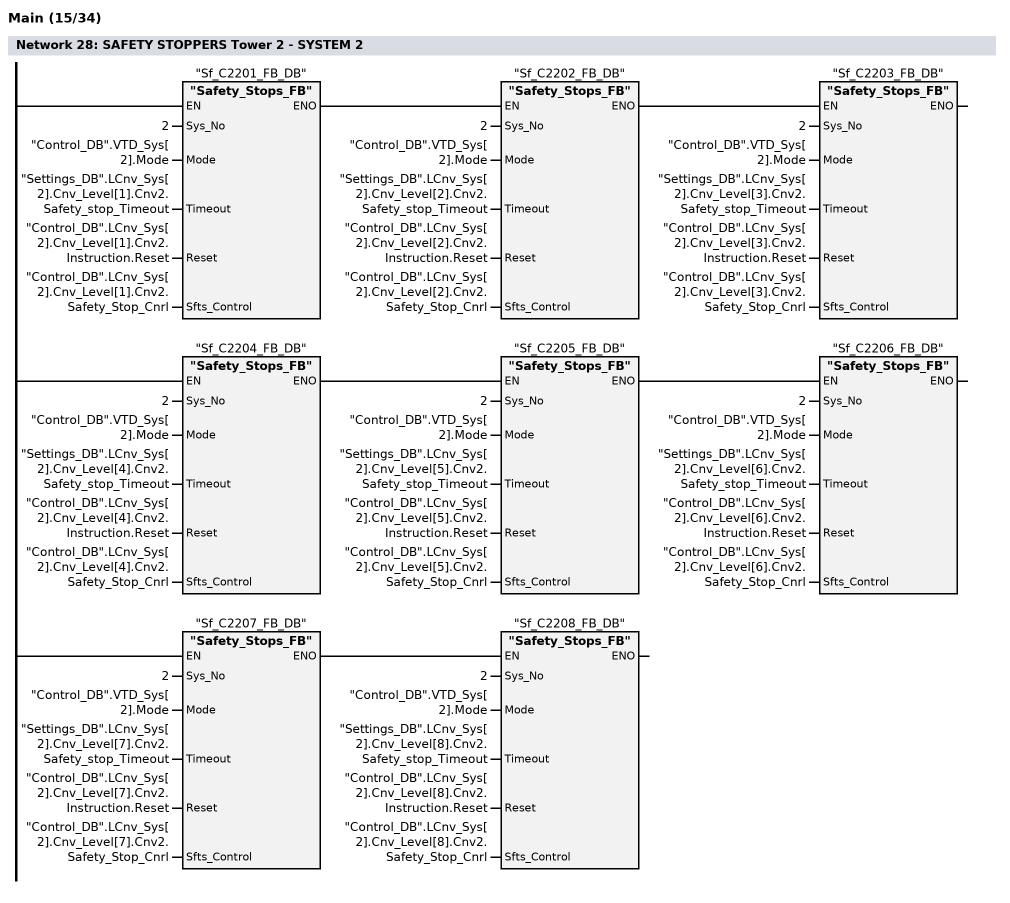
   RUNG wire#powerrail
      "Sf_C2201_FB_DB"(Sys_No := 2, Mode := "Control_DB".VTD_Sys[2].Mode, Timeout := "Settings_DB".LCnv_Sys[2].Cnv_Level[1].Cnv2.Safety_stop_Timeout, Reset := "Control_DB".LCnv_Sys[2].Cnv_Level[1].Cnv2.Instruction.Reset, Sfts_Control := "Control_DB".LCnv_Sys[2].Cnv_Level[1].Cnv2.Safety_Stop_Cnrl)
      "Sf_C2202_FB_DB"(Sys_No := 2, Mode := "Control_DB".VTD_Sys[2].Mode, Timeout := "Settings_DB".LCnv_Sys[2].Cnv_Level[2].Cnv2.Safety_stop_Timeout, Reset := "Control_DB".LCnv_Sys[2].Cnv_Level[2].Cnv2.Instruction.Reset, Sfts_Control := "Control_DB".LCnv_Sys[2].Cnv_Level[2].Cnv2.Safety_Stop_Cnrl)
      "Sf_C2203_FB_DB"(Sys_No := 2, Mode := "Control_DB".VTD_Sys[2].Mode, Timeout := "Settings_DB".LCnv_Sys[2].Cnv_Level[3].Cnv2.Safety_stop_Timeout, Reset := "Control_DB".LCnv_Sys[2].Cnv_Level[3].Cnv2.Instruction.Reset, Sfts_Control := "Control_DB".LCnv_Sys[2].Cnv_Level[3].Cnv2.Safety_Stop_Cnrl)
   END_RUNG
   RUNG wire#powerrail
      "Sf_C2204_FB_DB"(Sys_No := 2, Mode := "Control_DB".VTD_Sys[2].Mode, Timeout := "Settings_DB".LCnv_Sys[2].Cnv_Level[4].Cnv2.Safety_stop_Timeout, Reset := "Control_DB".LCnv_Sys[2].Cnv_Level[4].Cnv2.Instruction.Reset, Sfts_Control := "Control_DB".LCnv_Sys[2].Cnv_Level[4].Cnv2.Safety_Stop_Cnrl)
      "Sf_C2205_FB_DB"(Sys_No := 2, Mode := "Control_DB".VTD_Sys[2].Mode, Timeout := "Settings_DB".LCnv_Sys[2].Cnv_Level[5].Cnv2.Safety_stop_Timeout, Reset := "Control_DB".LCnv_Sys[2].Cnv_Level[5].Cnv2.Instruction.Reset, Sfts_Control := "Control_DB".LCnv_Sys[2].Cnv_Level[5].Cnv2.Safety_Stop_Cnrl)
      "Sf_C2206_FB_DB"(Sys_No := 2, Mode := "Control_DB".VTD_Sys[2].Mode, Timeout := "Settings_DB".LCnv_Sys[2].Cnv_Level[6].Cnv2.Safety_stop_Timeout, Reset := "Control_DB".LCnv_Sys[2].Cnv_Level[6].Cnv2.Instruction.Reset, Sfts_Control := "Control_DB".LCnv_Sys[2].Cnv_Level[6].Cnv2.Safety_Stop_Cnrl)
   END_RUNG
   RUNG wire#powerrail
      "Sf_C2207_FB_DB"(Sys_No := 2, Mode := "Control_DB".VTD_Sys[2].Mode, Timeout := "Settings_DB".LCnv_Sys[2].Cnv_Level[7].Cnv2.Safety_stop_Timeout, Reset := "Control_DB".LCnv_Sys[2].Cnv_Level[7].Cnv2.Instruction.Reset, Sfts_Control := "Control_DB".LCnv_Sys[2].Cnv_Level[7].Cnv2.Safety_Stop_Cnrl)
      "Sf_C2208_FB_DB"(Sys_No := 2, Mode := "Control_DB".VTD_Sys[2].Mode, Timeout := "Settings_DB".LCnv_Sys[2].Cnv_Level[8].Cnv2.Safety_stop_Timeout, Reset := "Control_DB".LCnv_Sys[2].Cnv_Level[8].Cnv2.Instruction.Reset, Sfts_Control := "Control_DB".LCnv_Sys[2].Cnv_Level[8].Cnv2.Safety_Stop_Cnrl)
   END_RUNG
   // the same network as SCL:
   "Sf_C2201_FB_DB"(Sys_No := 2,   // "Safety_Stops_FB"
                    Mode := "Control_DB".VTD_Sys[2].Mode,
                    Timeout := "Settings_DB".LCnv_Sys[2].Cnv_Level[1].Cnv2.Safety_stop_Timeout,
                    Reset := "Control_DB".LCnv_Sys[2].Cnv_Level[1].Cnv2.Instruction.Reset,
                    Sfts_Control := "Control_DB".LCnv_Sys[2].Cnv_Level[1].Cnv2.Safety_Stop_Cnrl,
                    ENO => #_w1);
   "Sf_C2202_FB_DB"(EN := #_w1,   // "Safety_Stops_FB"
                    Sys_No := 2,
                    Mode := "Control_DB".VTD_Sys[2].Mode,
                    Timeout := "Settings_DB".LCnv_Sys[2].Cnv_Level[2].Cnv2.Safety_stop_Timeout,
                    Reset := "Control_DB".LCnv_Sys[2].Cnv_Level[2].Cnv2.Instruction.Reset,
                    Sfts_Control := "Control_DB".LCnv_Sys[2].Cnv_Level[2].Cnv2.Safety_Stop_Cnrl,
                    ENO => #_w2);
   IF #_w2 THEN
       "Sf_C2203_FB_DB"(Sys_No := 2,   // "Safety_Stops_FB"
                        Mode := "Control_DB".VTD_Sys[2].Mode,
                        Timeout := "Settings_DB".LCnv_Sys[2].Cnv_Level[3].Cnv2.Safety_stop_Timeout,
                        Reset := "Control_DB".LCnv_Sys[2].Cnv_Level[3].Cnv2.Instruction.Reset,
                        Sfts_Control := "Control_DB".LCnv_Sys[2].Cnv_Level[3].Cnv2.Safety_Stop_Cnrl);
   END_IF;
   "Sf_C2204_FB_DB"(Sys_No := 2,   // "Safety_Stops_FB"
                    Mode := "Control_DB".VTD_Sys[2].Mode,
                    Timeout := "Settings_DB".LCnv_Sys[2].Cnv_Level[4].Cnv2.Safety_stop_Timeout,
                    Reset := "Control_DB".LCnv_Sys[2].Cnv_Level[4].Cnv2.Instruction.Reset,
                    Sfts_Control := "Control_DB".LCnv_Sys[2].Cnv_Level[4].Cnv2.Safety_Stop_Cnrl,
                    ENO => #_w3);
   "Sf_C2205_FB_DB"(EN := #_w3,   // "Safety_Stops_FB"
                    Sys_No := 2,
                    Mode := "Control_DB".VTD_Sys[2].Mode,
                    Timeout := "Settings_DB".LCnv_Sys[2].Cnv_Level[5].Cnv2.Safety_stop_Timeout,
                    Reset := "Control_DB".LCnv_Sys[2].Cnv_Level[5].Cnv2.Instruction.Reset,
                    Sfts_Control := "Control_DB".LCnv_Sys[2].Cnv_Level[5].Cnv2.Safety_Stop_Cnrl,
                    ENO => #_w4);
   IF #_w4 THEN
       "Sf_C2206_FB_DB"(Sys_No := 2,   // "Safety_Stops_FB"
                        Mode := "Control_DB".VTD_Sys[2].Mode,
                        Timeout := "Settings_DB".LCnv_Sys[2].Cnv_Level[6].Cnv2.Safety_stop_Timeout,
                        Reset := "Control_DB".LCnv_Sys[2].Cnv_Level[6].Cnv2.Instruction.Reset,
                        Sfts_Control := "Control_DB".LCnv_Sys[2].Cnv_Level[6].Cnv2.Safety_Stop_Cnrl);
   END_IF;
   "Sf_C2207_FB_DB"(Sys_No := 2,   // "Safety_Stops_FB"
                    Mode := "Control_DB".VTD_Sys[2].Mode,
                    Timeout := "Settings_DB".LCnv_Sys[2].Cnv_Level[7].Cnv2.Safety_stop_Timeout,
                    Reset := "Control_DB".LCnv_Sys[2].Cnv_Level[7].Cnv2.Instruction.Reset,
                    Sfts_Control := "Control_DB".LCnv_Sys[2].Cnv_Level[7].Cnv2.Safety_Stop_Cnrl,
                    ENO => #_w5);
   IF #_w5 THEN
       "Sf_C2208_FB_DB"(Sys_No := 2,   // "Safety_Stops_FB"
                        Mode := "Control_DB".VTD_Sys[2].Mode,
                        Timeout := "Settings_DB".LCnv_Sys[2].Cnv_Level[8].Cnv2.Safety_stop_Timeout,
                        Reset := "Control_DB".LCnv_Sys[2].Cnv_Level[8].Cnv2.Instruction.Reset,
                        Sfts_Control := "Control_DB".LCnv_Sys[2].Cnv_Level[8].Cnv2.Safety_Stop_Cnrl);
   END_IF;
END_REGION

REGION Network 29: SYSTEM 3
END_REGION

REGION Network 30: Level Conveyors Tower 1 - SYSTEM 3
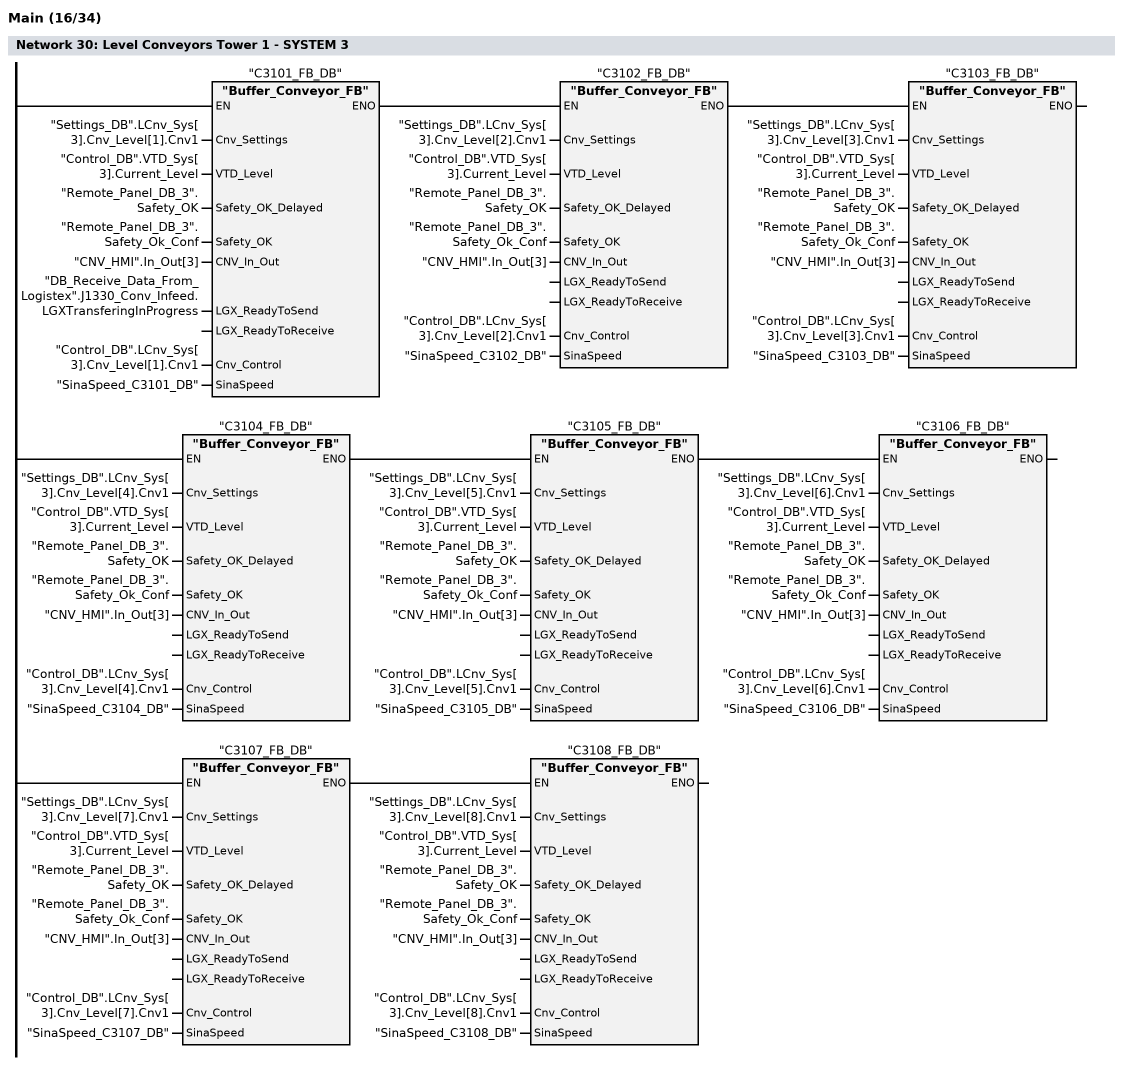
   RUNG wire#powerrail
      "C3101_FB_DB"(Cnv_Settings := "Settings_DB".LCnv_Sys[3].Cnv_Level[1].Cnv1, VTD_Level := "Control_DB".VTD_Sys[3].Current_Level, Safety_OK_Delayed := "Remote_Panel_DB_3".Safety_OK, Safety_OK := "Remote_Panel_DB_3".Safety_Ok_Conf, CNV_In_Out := "CNV_HMI".In_Out[3], LGX_ReadyToSend := "DB_Receive_Data_From_Logistex".J1330_Conv_Infeed.LGXTransferingInProgress, LGX_ReadyToReceive :=, Cnv_Control := "Control_DB".LCnv_Sys[3].Cnv_Level[1].Cnv1, SinaSpeed := "SinaSpeed_C3101_DB")
      "C3102_FB_DB"(Cnv_Settings := "Settings_DB".LCnv_Sys[3].Cnv_Level[2].Cnv1, VTD_Level := "Control_DB".VTD_Sys[3].Current_Level, Safety_OK_Delayed := "Remote_Panel_DB_3".Safety_OK, Safety_OK := "Remote_Panel_DB_3".Safety_Ok_Conf, CNV_In_Out := "CNV_HMI".In_Out[3], LGX_ReadyToSend :=, LGX_ReadyToReceive :=, Cnv_Control := "Control_DB".LCnv_Sys[3].Cnv_Level[2].Cnv1, SinaSpeed := "SinaSpeed_C3102_DB")
      "C3103_FB_DB"(Cnv_Settings := "Settings_DB".LCnv_Sys[3].Cnv_Level[3].Cnv1, VTD_Level := "Control_DB".VTD_Sys[3].Current_Level, Safety_OK_Delayed := "Remote_Panel_DB_3".Safety_OK, Safety_OK := "Remote_Panel_DB_3".Safety_Ok_Conf, CNV_In_Out := "CNV_HMI".In_Out[3], LGX_ReadyToSend :=, LGX_ReadyToReceive :=, Cnv_Control := "Control_DB".LCnv_Sys[3].Cnv_Level[3].Cnv1, SinaSpeed := "SinaSpeed_C3103_DB")
   END_RUNG
   RUNG wire#powerrail
      "C3104_FB_DB"(Cnv_Settings := "Settings_DB".LCnv_Sys[3].Cnv_Level[4].Cnv1, VTD_Level := "Control_DB".VTD_Sys[3].Current_Level, Safety_OK_Delayed := "Remote_Panel_DB_3".Safety_OK, Safety_OK := "Remote_Panel_DB_3".Safety_Ok_Conf, CNV_In_Out := "CNV_HMI".In_Out[3], LGX_ReadyToSend :=, LGX_ReadyToReceive :=, Cnv_Control := "Control_DB".LCnv_Sys[3].Cnv_Level[4].Cnv1, SinaSpeed := "SinaSpeed_C3104_DB")
      "C3105_FB_DB"(Cnv_Settings := "Settings_DB".LCnv_Sys[3].Cnv_Level[5].Cnv1, VTD_Level := "Control_DB".VTD_Sys[3].Current_Level, Safety_OK_Delayed := "Remote_Panel_DB_3".Safety_OK, Safety_OK := "Remote_Panel_DB_3".Safety_Ok_Conf, CNV_In_Out := "CNV_HMI".In_Out[3], LGX_ReadyToSend :=, LGX_ReadyToReceive :=, Cnv_Control := "Control_DB".LCnv_Sys[3].Cnv_Level[5].Cnv1, SinaSpeed := "SinaSpeed_C3105_DB")
      "C3106_FB_DB"(Cnv_Settings := "Settings_DB".LCnv_Sys[3].Cnv_Level[6].Cnv1, VTD_Level := "Control_DB".VTD_Sys[3].Current_Level, Safety_OK_Delayed := "Remote_Panel_DB_3".Safety_OK, Safety_OK := "Remote_Panel_DB_3".Safety_Ok_Conf, CNV_In_Out := "CNV_HMI".In_Out[3], LGX_ReadyToSend :=, LGX_ReadyToReceive :=, Cnv_Control := "Control_DB".LCnv_Sys[3].Cnv_Level[6].Cnv1, SinaSpeed := "SinaSpeed_C3106_DB")
   END_RUNG
   RUNG wire#powerrail
      "C3107_FB_DB"(Cnv_Settings := "Settings_DB".LCnv_Sys[3].Cnv_Level[7].Cnv1, VTD_Level := "Control_DB".VTD_Sys[3].Current_Level, Safety_OK_Delayed := "Remote_Panel_DB_3".Safety_OK, Safety_OK := "Remote_Panel_DB_3".Safety_Ok_Conf, CNV_In_Out := "CNV_HMI".In_Out[3], LGX_ReadyToSend :=, LGX_ReadyToReceive :=, Cnv_Control := "Control_DB".LCnv_Sys[3].Cnv_Level[7].Cnv1, SinaSpeed := "SinaSpeed_C3107_DB")
      "C3108_FB_DB"(Cnv_Settings := "Settings_DB".LCnv_Sys[3].Cnv_Level[8].Cnv1, VTD_Level := "Control_DB".VTD_Sys[3].Current_Level, Safety_OK_Delayed := "Remote_Panel_DB_3".Safety_OK, Safety_OK := "Remote_Panel_DB_3".Safety_Ok_Conf, CNV_In_Out := "CNV_HMI".In_Out[3], LGX_ReadyToSend :=, LGX_ReadyToReceive :=, Cnv_Control := "Control_DB".LCnv_Sys[3].Cnv_Level[8].Cnv1, SinaSpeed := "SinaSpeed_C3108_DB")
   END_RUNG
   // the same network as SCL:
   "C3101_FB_DB"(Cnv_Settings := "Settings_DB".LCnv_Sys[3].Cnv_Level[1].Cnv1,   // "Buffer_Conveyor_FB"
                 VTD_Level := "Control_DB".VTD_Sys[3].Current_Level,
                 Safety_OK_Delayed := "Remote_Panel_DB_3".Safety_OK,
                 Safety_OK := "Remote_Panel_DB_3".Safety_Ok_Conf,
                 CNV_In_Out := "CNV_HMI".In_Out[3],
                 LGX_ReadyToSend := "DB_Receive_Data_From_Logistex".J1330_Conv_Infeed.LGXTransferingInProgress,
                 Cnv_Control := "Control_DB".LCnv_Sys[3].Cnv_Level[1].Cnv1,
                 SinaSpeed := "SinaSpeed_C3101_DB",
                 ENO => #_w1);
   "C3102_FB_DB"(EN := #_w1,   // "Buffer_Conveyor_FB"
                 Cnv_Settings := "Settings_DB".LCnv_Sys[3].Cnv_Level[2].Cnv1,
                 VTD_Level := "Control_DB".VTD_Sys[3].Current_Level,
                 Safety_OK_Delayed := "Remote_Panel_DB_3".Safety_OK,
                 Safety_OK := "Remote_Panel_DB_3".Safety_Ok_Conf,
                 CNV_In_Out := "CNV_HMI".In_Out[3],
                 Cnv_Control := "Control_DB".LCnv_Sys[3].Cnv_Level[2].Cnv1,
                 SinaSpeed := "SinaSpeed_C3102_DB",
                 ENO => #_w2);
   IF #_w2 THEN
       "C3103_FB_DB"(Cnv_Settings := "Settings_DB".LCnv_Sys[3].Cnv_Level[3].Cnv1,   // "Buffer_Conveyor_FB"
                     VTD_Level := "Control_DB".VTD_Sys[3].Current_Level,
                     Safety_OK_Delayed := "Remote_Panel_DB_3".Safety_OK,
                     Safety_OK := "Remote_Panel_DB_3".Safety_Ok_Conf,
                     CNV_In_Out := "CNV_HMI".In_Out[3],
                     Cnv_Control := "Control_DB".LCnv_Sys[3].Cnv_Level[3].Cnv1,
                     SinaSpeed := "SinaSpeed_C3103_DB");
   END_IF;
   "C3104_FB_DB"(Cnv_Settings := "Settings_DB".LCnv_Sys[3].Cnv_Level[4].Cnv1,   // "Buffer_Conveyor_FB"
                 VTD_Level := "Control_DB".VTD_Sys[3].Current_Level,
                 Safety_OK_Delayed := "Remote_Panel_DB_3".Safety_OK,
                 Safety_OK := "Remote_Panel_DB_3".Safety_Ok_Conf,
                 CNV_In_Out := "CNV_HMI".In_Out[3],
                 Cnv_Control := "Control_DB".LCnv_Sys[3].Cnv_Level[4].Cnv1,
                 SinaSpeed := "SinaSpeed_C3104_DB",
                 ENO => #_w3);
   "C3105_FB_DB"(EN := #_w3,   // "Buffer_Conveyor_FB"
                 Cnv_Settings := "Settings_DB".LCnv_Sys[3].Cnv_Level[5].Cnv1,
                 VTD_Level := "Control_DB".VTD_Sys[3].Current_Level,
                 Safety_OK_Delayed := "Remote_Panel_DB_3".Safety_OK,
                 Safety_OK := "Remote_Panel_DB_3".Safety_Ok_Conf,
                 CNV_In_Out := "CNV_HMI".In_Out[3],
                 Cnv_Control := "Control_DB".LCnv_Sys[3].Cnv_Level[5].Cnv1,
                 SinaSpeed := "SinaSpeed_C3105_DB",
                 ENO => #_w4);
   IF #_w4 THEN
       "C3106_FB_DB"(Cnv_Settings := "Settings_DB".LCnv_Sys[3].Cnv_Level[6].Cnv1,   // "Buffer_Conveyor_FB"
                     VTD_Level := "Control_DB".VTD_Sys[3].Current_Level,
                     Safety_OK_Delayed := "Remote_Panel_DB_3".Safety_OK,
                     Safety_OK := "Remote_Panel_DB_3".Safety_Ok_Conf,
                     CNV_In_Out := "CNV_HMI".In_Out[3],
                     Cnv_Control := "Control_DB".LCnv_Sys[3].Cnv_Level[6].Cnv1,
                     SinaSpeed := "SinaSpeed_C3106_DB");
   END_IF;
   "C3107_FB_DB"(Cnv_Settings := "Settings_DB".LCnv_Sys[3].Cnv_Level[7].Cnv1,   // "Buffer_Conveyor_FB"
                 VTD_Level := "Control_DB".VTD_Sys[3].Current_Level,
                 Safety_OK_Delayed := "Remote_Panel_DB_3".Safety_OK,
                 Safety_OK := "Remote_Panel_DB_3".Safety_Ok_Conf,
                 CNV_In_Out := "CNV_HMI".In_Out[3],
                 Cnv_Control := "Control_DB".LCnv_Sys[3].Cnv_Level[7].Cnv1,
                 SinaSpeed := "SinaSpeed_C3107_DB",
                 ENO => #_w5);
   IF #_w5 THEN
       "C3108_FB_DB"(Cnv_Settings := "Settings_DB".LCnv_Sys[3].Cnv_Level[8].Cnv1,   // "Buffer_Conveyor_FB"
                     VTD_Level := "Control_DB".VTD_Sys[3].Current_Level,
                     Safety_OK_Delayed := "Remote_Panel_DB_3".Safety_OK,
                     Safety_OK := "Remote_Panel_DB_3".Safety_Ok_Conf,
                     CNV_In_Out := "CNV_HMI".In_Out[3],
                     Cnv_Control := "Control_DB".LCnv_Sys[3].Cnv_Level[8].Cnv1,
                     SinaSpeed := "SinaSpeed_C3108_DB");
   END_IF;
END_REGION

